// §3.8b — "restore is fail-closed and never silent". Every module that ran
// M_RestoreStationCfg and found an unrecognized image is holding one report;
// this takes them and annunciates each with the OWNING module's canonical path,
// which is what makes the message actionable instead of "something was lost".
//
// The event is AUTO_RESET and therefore never blocking: the consequence belongs
// to E_ConfigRestorePolicy, evaluated in ReleaseReportStart, so a station that
// declared DEFAULTS_AND_ANNUNCIATE really does run while the annunciation
// stands. It stays open until an ENGINEER acknowledges it, because nothing
// makes a lost image come back and an event that closed itself would be a lie.
METHOD PRIVATE _M_DrainRestoreLoss
VAR
    guard    : INT;
    path     : STRING(80);
    expected : UINT;
    found    : UINT;
END_VAR
// §7.7(c) - the local user table is retained outside the module walk; its loss
// is announced and acknowledged exactly like a module's.
IF Access.M_TakeRestoreLoss() THEN
    path := CONCAT(_name, '.Access');
    _M_AnnounceRestoreLoss(Path := path, Text := 'std.error.accessRestoreLost');
END_IF
// Bounded per scan (§5.6): losses are one-shot, so a large subtree simply
// finishes draining over the next few scans instead of stretching one.
FOR guard := 1 TO PL_Fraktal.MAX_EM_CHILDREN DO
    IF NOT M_TakeRestoreLoss(Path => path, Expected => expected, Found => found) THEN
        RETURN;
    END_IF
    _M_AnnounceRestoreLoss(Path := path, Text := 'std.error.configRestoreLost');
END_FOR
END_METHOD

// §3.8b - publish one lost image and open (or extend) its annunciation.
METHOD PRIVATE _M_AnnounceRestoreLoss
VAR_INPUT
    Path : STRING(80);
    Text : STRING(80);
END_VAR
ConfigPersist.RestoreLost := TRUE;
ConfigPersist.RestoreAcknowledged := FALSE;
ConfigPersist.LostPath := Path;
IF _restoreEvt = 0 THEN
    _restoreEvt := AlarmLog.Raise(Reason := E_Reason.CONFIG_RESTORE_LOST,
        Text := Text, Source := Path,
        Severity := E_Severity.MED, Category := E_Category.SYSTEM,
        ResetClass := E_ResetClass.AUTO_RESET);
ELSE
    // A second losing owner gets its own ring entry: a summary that named only
    // the first would hide the rest of the damage.
    _M_RaiseMaintenance(Reason := E_Reason.CONFIG_RESTORE_LOST, Text := Text);
END_IF
END_METHOD

// §3.8b — an operator of at least ENGINEER level accepts that a configuration
// image was lost. Under BLOCK_UNTIL_ACKNOWLEDGED this is what releases
// START_STOP again; under DEFAULTS_AND_ANNUNCIATE it is what clears the
// standing annunciation.
//
// The level is checked directly rather than through a gated action, because
// §3.8b names ENGINEER specifically and a station may legitimately have left
// DATA_WRITE or CONFIG_SET open to a lower level. Acknowledging a lost
// commissioning is a different decision from editing a value.
METHOD AcknowledgeConfigRestore : BOOL
AcknowledgeConfigRestore := FALSE;
IF Access.CurrentLevel < E_AccessLevel.ENGINEER THEN
    RETURN;
END_IF
IF NOT ConfigPersist.RestoreLost THEN
    RETURN;                                // nothing to acknowledge
END_IF
ConfigPersist.RestoreAcknowledged := TRUE;
IF _restoreEvt > 0 THEN
    AlarmLog.Gone(Slot := _restoreEvt);
    _restoreEvt := 0;
END_IF
Access.RecordActivity();
AcknowledgeConfigRestore := TRUE;
END_METHOD

// §3.8b — refuse a set operation, naming the offending record. "One rejection
// aborts the whole load naming the offending (Scope, WriteKey)": a refusal that
// says only "rejected" leaves an engineer diffing two machines by hand.
METHOD PRIVATE _M_RejectConfigSet
VAR_INPUT
    Scope : STRING(80);
    Key   : STRING(160);
END_VAR
ConfigPersist.LastRejectScope := Scope;
ConfigPersist.LastRejectKey := Key;
_M_RaiseMaintenance(Reason := E_Reason.CONFIG_SET_REJECTED,
    Text := 'std.error.configSetRejected');
END_METHOD

// §3.8b — the gate every set operation shares: CONFIG_SET (never DATA_WRITE —
// replacing a machine's entire parametrization is not the same decision as
// changing one number), a wired store, and the owning root READY.
METHOD PRIVATE _M_SetOpAllowed : BOOL
_M_SetOpAllowed := FALSE;
IF NOT _M_ConfigRestored() THEN
    RETURN;
END_IF
IF NOT Access.PermitsLogged(Gate := E_GatedAction.CONFIG_SET) THEN
    RETURN;
END_IF
IF _configStore = 0 THEN
    RETURN;
END_IF
IF _exec <> E_ExecState.READY THEN
    RETURN;
END_IF
_M_SetOpAllowed := TRUE;
END_METHOD

// §3.8b - remove a named set. Gated exactly like save and load (CONFIG_SET, a
// wired store, the root READY) because removing somebody's commissioned set is
// the same order of decision as replacing it, and audited with the set name.
// A store that has held MAX_CONFIG_SETS names needs this to hold a new one.
METHOD DeleteConfigSet : BOOL
VAR_INPUT
    SetName : STRING(80);
END_VAR
DeleteConfigSet := FALSE;
ConfigPersist.LastSetName := SetName;
ConfigPersist.LastSetRecords := 0;
IF NOT _M_SetOpAllowed() THEN
    RETURN;
END_IF
IF NOT _configStore.M_Delete(SetName := SetName) THEN
    RETURN;
END_IF
DeleteConfigSet := TRUE;
// The store's retained memory changed; not durable until written out.
_M_MarkPersistPending();
ListConfigSets();                          // the published listing follows
END_METHOD

// §3.8d - the effective level to read or write one registered value, from
// what its owning module declared and this root's policy. The root's own
// framework keys (unit.modePolicy.*) are in the built-in class. An unknown key
// resolves to ADMIN: the write path refuses it anyway, and a level check must
// never be the thing that lets an unknown key through.
METHOD PRIVATE _M_DataLevelOf : E_AccessLevel
VAR_INPUT
    TargetPath : STRING(255);
    WriteKey   : STRING(160);
    ForWrite   : BOOL;
END_VAR
VAR
    grant    : ST_ConfigAccess;
    minLevel : E_AccessLevel;
END_VAR
_M_DataLevelOf := E_AccessLevel.ADMIN;
IF (TargetPath = Status.Name) AND (LEFT(WriteKey, 16) = 'unit.modePolicy.') THEN
    _M_DataLevelOf := Access.M_DataLevel(ClassId := '', MinLevel := E_AccessLevel.NONE,
        ForWrite := ForWrite);
    RETURN;
END_IF
IF NOT M_ConfigAccessOf(Scope := TargetPath, WriteKey := WriteKey, Grant := grant) THEN
    RETURN;
END_IF
IF ForWrite THEN
    minLevel := grant.MinWriteLevel;
ELSE
    minLevel := grant.MinReadLevel;
END_IF
_M_DataLevelOf := Access.M_DataLevel(ClassId := grant.ClassId, MinLevel := minLevel,
    ForWrite := ForWrite);
END_METHOD

// §3.8d - declare a project data class on this root, at Setup. The levels are
// defaults: a class the deployment already edited keeps its persisted levels.
METHOD M_DeclareDataClass : BOOL
VAR_INPUT
    ClassId    : STRING(80);
    LabelKey   : STRING(160);
    ReadLevel  : E_AccessLevel;
    WriteLevel : E_AccessLevel;
END_VAR
M_DeclareDataClass := Access.M_DeclareClass(ClassId := ClassId,
    LabelKey := LabelKey, ReadLevel := ReadLevel, WriteLevel := WriteLevel);
END_METHOD

// §3.8d/§7.7(b) - edit a class's read or write level. The same gate as
// every other policy edit (ACCESS_POLICY), audited through the mailbox.
METHOD SetDataClassLevel : BOOL
VAR_INPUT
    ClassId  : STRING(160);
    Level    : DINT;
    ForWrite : BOOL;
END_VAR
VAR
    levelReq : E_AccessLevel;
END_VAR
SetDataClassLevel := FALSE;
IF NOT Access.PermitsLogged(Gate := E_GatedAction.ACCESS_POLICY) THEN
    RETURN;
END_IF
IF (Level < TO_DINT(E_AccessLevel.NONE)) OR (Level > TO_DINT(E_AccessLevel.ADMIN))
OR (LEN(ClassId) > 40) THEN
    RETURN;
END_IF
levelReq := Level;                          // range-checked above
SetDataClassLevel := Access.M_SetClassLevel(ClassId := ClassId,
    Level := levelReq, ForWrite := ForWrite);
IF SetDataClassLevel THEN
    ConfigRev := ConfigRev + 1;             // every manifest level may have moved
END_IF
END_METHOD

// §3.8e - TRUE when a (Scope, WriteKey) the subtree did not own names a value of
// the line this Unit references: the line is published under this Unit's own
// scope, and its keys alone begin 'line.'.
METHOD PRIVATE _M_IsLineKey : BOOL
VAR_INPUT
    Scope    : STRING(255);
    WriteKey : STRING(160);
END_VAR
_M_IsLineKey := (_pLine <> 0) AND (Scope = Status.Name)
    AND (LEFT(WriteKey, 5) = 'line.');
END_METHOD

// §3.8e - the subtree first; a line key it does not own goes to the line.
METHOD M_ApplyConfigWrite : BOOL
VAR_INPUT
    Scope     : STRING(255);
    WriteKey  : STRING(160);
    Revision  : UDINT;
    TextValue : STRING(255);
    RootReady : BOOL;
END_VAR
M_ApplyConfigWrite := SUPER^.M_ApplyConfigWrite(Scope := Scope,
    WriteKey := WriteKey, Revision := Revision, TextValue := TextValue,
    RootReady := RootReady);
IF (NOT M_ApplyConfigWrite) AND _M_IsLineKey(Scope := Scope, WriteKey := WriteKey) THEN
    M_ApplyConfigWrite := _pLine^.M_ApplyConfigWrite(Scope := _pLine^.Status.Name,
        WriteKey := WriteKey, Revision := Revision, TextValue := TextValue,
        RootReady := RootReady);
END_IF
END_METHOD

// §3.8e - the staging walk is the write walk, line leg included.
METHOD M_StageConfigWrite : BOOL
VAR_INPUT
    Scope     : STRING(255);
    WriteKey  : STRING(160);
    Revision  : UDINT;
    TextValue : STRING(255);
    RootReady : BOOL;
END_VAR
M_StageConfigWrite := SUPER^.M_StageConfigWrite(Scope := Scope,
    WriteKey := WriteKey, Revision := Revision, TextValue := TextValue,
    RootReady := RootReady);
IF (NOT M_StageConfigWrite) AND _M_IsLineKey(Scope := Scope, WriteKey := WriteKey) THEN
    M_StageConfigWrite := _pLine^.M_StageConfigWrite(Scope := _pLine^.Status.Name,
        WriteKey := WriteKey, Revision := Revision, TextValue := TextValue,
        RootReady := RootReady);
END_IF
END_METHOD

// §3.8e - the capture walk is the write walk, line leg included.
METHOD M_ApplyCapture : BOOL
VAR_INPUT
    Scope     : STRING(255);
    WriteKey  : STRING(160);
    Revision  : UDINT;
    RootReady : BOOL;
END_VAR
M_ApplyCapture := SUPER^.M_ApplyCapture(Scope := Scope, WriteKey := WriteKey,
    Revision := Revision, RootReady := RootReady);
IF (NOT M_ApplyCapture) AND _M_IsLineKey(Scope := Scope, WriteKey := WriteKey) THEN
    M_ApplyCapture := _pLine^.M_ApplyCapture(Scope := _pLine^.Status.Name,
        WriteKey := WriteKey, Revision := Revision, RootReady := RootReady);
END_IF
END_METHOD

// §3.8e/§3.8d - the access walk is the write walk, line leg included, so a line
// value is checked against the level the line declared for it.
METHOD M_ConfigAccessOf : BOOL
VAR_INPUT
    Scope    : STRING(255);
    WriteKey : STRING(160);
END_VAR
VAR_IN_OUT
    Grant : ST_ConfigAccess;
END_VAR
M_ConfigAccessOf := SUPER^.M_ConfigAccessOf(Scope := Scope, WriteKey := WriteKey,
    Grant := Grant);
IF (NOT M_ConfigAccessOf) AND _M_IsLineKey(Scope := Scope, WriteKey := WriteKey) THEN
    M_ConfigAccessOf := _pLine^.M_ConfigAccessOf(Scope := _pLine^.Status.Name,
        WriteKey := WriteKey, Grant := Grant);
END_IF
END_METHOD

// Core §3.8a - declare this root's own recipe record (its ParCfg) and the
// provider it is loaded from. The PAR_CFG values registered inside it become
// editable for EVERY model the root offers (AvailableModels), not only the
// active one, and an edit is written back to the provider's record so a
// changeover keeps it - when the provider is also an I_RecipeStore.
METHOD M_RegisterModelData : BOOL
VAR_INPUT
    pData     : PVOID;
    Size      : UDINT;
    RecipeKey : STRING(80);
    Provider  : I_RecipeProvider;
END_VAR
M_RegisterModelData := FALSE;
IF (pData = 0) OR (Size = 0) OR (Size > PL_Fraktal.MAX_MODEL_DATA_BYTES)
OR (RecipeKey = '') OR (Provider = 0) THEN
    RETURN;
END_IF
_modelProvider := Provider;
__QUERYINTERFACE(Provider, _modelCatalog);
_modelKey := RecipeKey;
M_RegisterModelData := _M_SetModelRegion(pRegion := pData, Size := Size);
END_METHOD

// Serve model-scoped values of AvailableModels[Index] for this one request. 0,
// or the active model's index, is the live record and opens nothing. The record
// is loaded over a copy of the live one, so the provider's SchemaVersion check
// compares like with like. FALSE = no such model, or its record did not load.
METHOD PRIVATE _M_OpenModelView : BOOL
VAR_INPUT
    Index : UDINT;
END_VAR
_M_OpenModelView := FALSE;
_pModelView := 0;
_viewModelCode := '';
IF Index = 0 THEN
    _M_OpenModelView := TRUE;
    RETURN;
END_IF
IF (_modelProvider = 0) OR (_pModelRegion = 0)
OR (Index > TO_UDINT(AvailableModelCount)) THEN
    RETURN;
END_IF
IF AvailableModels[Index].ModelCode = Model.ModelCode THEN
    _M_OpenModelView := TRUE;              // the active model: its record is live
    RETURN;
END_IF
MEMCPY(destAddr := ADR(_modelBuf), srcAddr := _pModelRegion, n := _modelRegionSize);
IF NOT _modelProvider.Load(ModelCode := AvailableModels[Index].ModelCode,
        RecipeKey := _modelKey, pParCfg := ADR(_modelBuf), Size := _modelRegionSize) THEN
    RETURN;
END_IF
_viewModelCode := AvailableModels[Index].ModelCode;
_pModelView := ADR(_modelBuf);
_M_OpenModelView := TRUE;
END_METHOD

// §3.8a - WriteConfig for the model AvailableModels[ModelIndex] (0 = the active
// model). A model-data value is stored in that model's record and saved back to
// the provider; any other value is written as WriteConfig writes it.
METHOD WriteModelConfig : BOOL
VAR_INPUT
    ModelIndex : UDINT;
    TargetPath : STRING(255);
    WriteKey   : STRING(160);
    Revision   : DINT;
    TextValue  : STRING(255);
END_VAR
WriteModelConfig := FALSE;
IF NOT _M_OpenModelView(Index := ModelIndex) THEN
    RETURN;
END_IF
WriteModelConfig := WriteConfig(TargetPath := TargetPath, WriteKey := WriteKey,
    Revision := Revision, TextValue := TextValue);
_pModelView := 0;
END_METHOD

// §3.8a - the manifest walk (M_AppendConfig) with the model-data values of
// AvailableModels[ModelIndex] (0 = the active model). FALSE = no such model.
// For another model the walk yields that model's data only: the rest of the
// manifest is the running station's and is served by index 0.
METHOD M_AppendModelConfig : BOOL
VAR_INPUT
    Pager      : REFERENCE TO FB_ConfigPager;
    ModelIndex : UDINT;
END_VAR
M_AppendModelConfig := FALSE;
IF NOT _M_OpenModelView(Index := ModelIndex) THEN
    RETURN;
END_IF
Pager.M_SetModelOnly(Enabled := ModelIndex > 0);
M_AppendConfig(Pager := Pager);
Pager.M_SetModelOnly(Enabled := FALSE);
_pModelView := 0;
M_AppendModelConfig := TRUE;
END_METHOD

// Write the record a model-scoped value was just stored into back to the
// provider: the viewed model's buffer, or the live record for the active model.
METHOD PRIVATE _M_SaveModelData : BOOL
VAR
    store : I_RecipeStore;
END_VAR
_M_SaveModelData := FALSE;
IF _modelProvider = 0 THEN
    RETURN;
END_IF
IF NOT __QUERYINTERFACE(_modelProvider, store) THEN
    RETURN;
END_IF
IF _pModelView <> 0 THEN
    _M_SaveModelData := store.Save(ModelCode := _viewModelCode, RecipeKey := _modelKey,
        pData := _pModelView, Size := _modelRegionSize);
ELSE
    _M_SaveModelData := store.Save(ModelCode := Model.ModelCode, RecipeKey := _modelKey,
        pData := _pModelRegion, Size := _modelRegionSize);
END_IF
END_METHOD

// §3.8e/§8.5.2 - reference the line this root belongs to (owner or mirror, on
// this controller). A Unit references at most one line; 0 detaches it.
METHOD SetLine : BOOL
VAR_INPUT
    pLine : POINTER TO FB_LineData;
END_VAR
_pLine := pLine;
_lineHost := FALSE;
IF pLine <> 0 THEN
    // The first root to reference a line hosts it (ticks it, lends its log); a
    // line is never a child, so nothing else would run it (§3.8e(a)).
    _lineHost := pLine^.M_BindHost(pHost := THIS, pAlarmLog := ADR(AlarmLog));
END_IF
_shiftInit := FALSE;
CurrentShift := 0;
SetLine := (pLine <> 0);
END_METHOD

// Evaluate only at a finite boundary, or after an empty-calendar edit.
METHOD M_ShiftTick : BOOL
VAR_INPUT
    Now : DT;
    Synchronized : BOOL;
END_VAR
VAR
    idx : INT;
    started : DT;
    ending : DT;
    target : UDINT;
    crossed : BOOL;
    quality : BOOL;
END_VAR
M_ShiftTick := FALSE;
IF _pLine = 0 THEN CurrentShift := 0; ShiftProductionTarget := 0; RETURN; END_IF
IF _shiftInit THEN
    IF Now < _shiftLastNow THEN _shiftSync := FALSE; END_IF
    _shiftLastNow := Now;
    IF (_shiftEnd <> DT#1970-01-01-00:00:00) AND (Now < _shiftEnd) THEN RETURN; END_IF
    IF Now < ShiftStartedAt THEN RETURN; END_IF // no negative history after a backward jump
    IF (_shiftEnd = DT#1970-01-01-00:00:00)
    AND (_shiftCalendarRev = _pLine^.OutImm.Revision) THEN RETURN; END_IF
END_IF
IF NOT _pLine^.M_ShiftInterval(Now := Now, ShiftIndex => idx,
        StartAt => started, EndAt => ending, Target => target) THEN
    _shiftSync := FALSE; RETURN;
END_IF
crossed := _shiftInit AND (_shiftEnd <> DT#1970-01-01-00:00:00);
IF _shiftInit AND NOT crossed AND (idx = 0) THEN
    // Empty/off interval continues; an edit must not erase accrued production.
    _shiftEnd := ending;
    _shiftCalendarRev := _pLine^.OutImm.Revision;
    RETURN;
END_IF
IF _shiftInit THEN
    quality := Synchronized;
    IF crossed AND (DT_TO_UDINT(Now) > DT_TO_UDINT(_shiftEnd) + 1) THEN quality := FALSE; END_IF
    _M_CloseShift(Now := Now, Synchronized := quality);
    M_ShiftTick := TRUE;
END_IF
_shiftInit := TRUE;
CurrentShift := idx;
ShiftStartedAt := Now; // observed start, never invent production before attachment/jump
ShiftProductionTarget := target;
_shiftEnd := ending;
_shiftLastNow := Now;
_shiftCalendarRev := _pLine^.OutImm.Revision;
_shiftSync := Synchronized;
_shiftManualReset := FALSE;
END_METHOD

// §8.5.2(b) - one operation in one scan: record the ending shift as its figures stood,
// then reset the per-shift counts and OEE accumulators (the trend ring is kept). A
// boundary on an unsynchronized clock still closes - stopping the accounting would
// lose more than a late boundary does - and the record says so.
METHOD PRIVATE _M_CloseShift
VAR_INPUT
    Now          : DT;
    Synchronized : BOOL;
END_VAR
VAR
    i         : INT;
    auditSlot : INT;
END_VAR
_M_OeeCompute(); // capture current factors before counters are cleared
FOR i := PL_Fraktal.MAX_SHIFT_HISTORY TO 2 BY -1 DO
    ShiftHistory[i] := ShiftHistory[i - 1];
END_FOR
IF ShiftHistoryCount >= PL_Fraktal.MAX_SHIFT_HISTORY THEN
    ShiftHistoryTruncated := TRUE;
ELSE
    ShiftHistoryCount := ShiftHistoryCount + 1;
END_IF
ShiftHistory[1].SchemaVersion := 3;
ShiftHistory[1].ProductionTarget := ShiftProductionTarget;
ShiftHistory[1].ShiftIndex := CurrentShift;
ShiftHistory[1].StartAt := ShiftStartedAt;
ShiftHistory[1].EndAt := Now;
ShiftHistory[1].TimeSynchronized := _shiftSync AND Synchronized;
ShiftHistory[1].ManualReset := _shiftManualReset;
ShiftHistory[1].GoodCount := GoodCount;
ShiftHistory[1].NokCount := NokCount;
ShiftHistory[1].ReworkCount := ReworkCount;
ShiftHistory[1].RunMs := Oee.RunMs;
ShiftHistory[1].DownMs := Oee.DownMs;
ShiftHistory[1].IdleMs := Oee.IdleMs;
ShiftHistory[1].Availability := Oee.Availability;
ShiftHistory[1].AvailValid := Oee.AvailValid;
ShiftHistory[1].Performance := Oee.Performance;
ShiftHistory[1].PerfValid := Oee.PerfValid;
ShiftHistory[1].Quality := Oee.Quality;
ShiftHistory[1].QualValid := Oee.QualValid;
ShiftHistory[1].Oee := Oee.Oee;
ShiftHistory[1].OeeValid := Oee.OeeValid;
_oeeGoodBase := 0;
_oeeNokBase := 0;
GoodCount := 0;
NokCount := 0;
ReworkCount := 0;
Oee.RunMs := 0;
Oee.DownMs := 0;
Oee.IdleMs := 0;
_M_OeeCompute();
auditSlot := AlarmLog.Raise(Reason := E_Reason.NONE, Text := 'std.audit.shiftClosed',
    Source := _name, Severity := E_Severity.LOW, Category := E_Category.SYSTEM,
    ResetClass := E_ResetClass.AUTO_RESET);
IF auditSlot > 0 THEN
    AlarmLog.Gone(Slot := auditSlot);    // come+gone: into the ring and the event sink
END_IF
END_METHOD

// §3.8b — save the current parametrization as a named set.
//
// The set is a PROJECTION of the same deterministic walk that builds the
// §3.10.2 manifest: M_AppendConfig runs exactly as a QUERY_CONFIG would run it,
// and the pager files every capability of the requested ConfigKind as a
// (Scope, WriteKey) record. There is no second enumeration of "what this
// station's configuration consists of" to drift from the first (§1.1 O9).
//
// Kind selects which of the two kinds of set this is: STATION_CFG for a station
// set (deployment data), PAR_CFG for a model set (one model's recipe data).
METHOD SaveConfigSet : BOOL
VAR_INPUT
    SetName : STRING(80);
    Kind    : E_ConfigKind;
END_VAR
VAR
    info    : ST_ConfigSetInfo;
    records : INT;
END_VAR
SaveConfigSet := FALSE;
ConfigPersist.LastSetName := SetName;
ConfigPersist.LastSetRecords := 0;
IF NOT _M_SetOpAllowed() THEN
    RETURN;
END_IF
IF SetName = '' THEN
    RETURN;
END_IF
info.Used := TRUE;
info.SetName := SetName;
info.RootIdentity := Status.Name;
info.SetSchema := CONFIG_SET_SCHEMA;
info.ConfigRev := ConfigRev;
info.Kind := Kind;
IF Kind = E_ConfigKind.PAR_CFG THEN
    info.ModelCode := Model.ModelCode;     // a model set belongs to ONE model
ELSE
    info.ModelCode := '';
END_IF
info.RecordCount := 0;
info.CreatedAt := F_Now();
info.TimeSynchronized := F_TimeSynchronized();
IF NOT _configPager.M_SetupSetSave(Store := _configStore, Info := info) THEN
    RETURN;
END_IF
M_AppendConfig(Pager := _configPager);     // the SAME walk as the manifest
SaveConfigSet := _configPager.M_FinishSetSave(Records => records);
ConfigPersist.LastSetRecords := records;
IF SaveConfigSet THEN
    // The set now lives in the store's retained memory, which is not durable
    // until it is written out - the same promise as any other accepted write.
    _M_MarkPersistPending();
END_IF
END_METHOD

// §3.8b — apply a named set. STAGED and ALL-OR-NOTHING.
//
// Pass 1 validates every record through its owning module's typed handler and
// changes nothing. Only if all of them pass does pass 2 apply them. A
// half-applied machine parametrization is never a valid outcome, and the only
// way to guarantee that is to know the answer for every record before touching
// the first one.
//
// A record whose capability no longer exists fails pass 1 like any other and is
// REPORTED by name - never silently dropped, because a set that quietly skipped
// the one value that mattered restores a machine to almost its commissioned
// state, which is the failure that is hardest to notice.
METHOD LoadConfigSet : BOOL
VAR_INPUT
    SetName : STRING(80);
END_VAR
VAR
    info    : ST_ConfigSetInfo;
END_VAR
LoadConfigSet := FALSE;
ConfigPersist.LastSetName := SetName;
ConfigPersist.LastSetRecords := 0;
ConfigPersist.LastRejectScope := '';
ConfigPersist.LastRejectKey := '';
IF NOT _M_SetOpAllowed() THEN
    RETURN;
END_IF
IF NOT _M_CopySet(SetName := SetName) THEN
    RETURN;
END_IF
IF NOT _loadSnapshot.M_ReadInfo(SetName := SetName, Info := info) THEN
    _M_RejectConfigSet(Scope := '', Key := SetName);
    RETURN;
END_IF
IF info.RootIdentity <> Status.Name THEN
    // The set carries the identity of the root that produced it precisely so
    // this can be asked. Every record's Scope is prefixed by that identity, so
    // a mismatch would fail record by record anyway - naming the root instead
    // tells the operator WHY in one line.
    _M_RejectConfigSet(Scope := info.RootIdentity, Key := '');
    RETURN;
END_IF
IF info.Kind = E_ConfigKind.PAR_CFG THEN
    // §3.8b: a MODEL set "shall be applied through the §3.8 changeover
    // transaction (PrepareRecipe -> recursive readiness -> infallible
    // CommitRecipe), never as a sequence of per-field writes". Applying it here
    // would be exactly that forbidden sequence, so it is refused. Saving a
    // model set is supported; loading one is a changeover this build does not
    // implement, and refusing is the honest half of that.
    _M_RejectConfigSet(Scope := info.ModelCode, Key := '');
    RETURN;
END_IF
IF NOT _M_CaptureConfig(SetName := '_validation', Kind := info.Kind, ModelIndex := 0) THEN RETURN; END_IF
IF NOT _M_ValidateSetShape(Store := _loadSnapshot, Info := info, AnyRevision := FALSE) THEN
    RETURN;
END_IF
IF NOT _M_ApplySet(SetName := SetName, RecordCount := info.RecordCount, Kind := info.Kind,
        Restoring := FALSE) THEN
    RETURN;
END_IF
ConfigRev := ConfigRev + 1;
ConfigPersist.LastSetRecords := info.RecordCount;
_M_MarkPersistPending();
_M_RaiseMaintenance(Reason := E_Reason.EVENT_CONFIG_SET_APPLIED,
    Text := 'std.audit.configSetApplied');
LoadConfigSet := TRUE;
END_METHOD

// §3.8b - replay the set frozen in _loadSnapshot. STAGED and ALL-OR-NOTHING:
// pass 1 validates every record through its owning module's typed handler and
// changes nothing; only if all of them pass does pass 2 apply them. A record
// whose capability no longer exists fails pass 1 like any other and is named.
//
// Shared by an operator's LoadConfigSet and the start-up restore of the live
// documents. Restoring skips the session's per-value level (§3.8d(e)): those
// values were accepted once already, and replaying them is the machine's act,
// not an operator's. With a model view open the values go to that record.
METHOD PRIVATE _M_ApplySet : BOOL
VAR_INPUT
    SetName     : STRING(80);
    RecordCount : INT;
    Kind        : E_ConfigKind;
    Restoring   : BOOL;
END_VAR
VAR
    record    : ST_ConfigRecord;
    i         : INT;
    applied   : BOOL;
    lineBatch : BOOL;
END_VAR
_M_ApplySet := FALSE;
lineBatch := (Kind = E_ConfigKind.LINE_CFG) AND (_pLine <> 0);
IF lineBatch THEN
    IF NOT _pLine^.M_BeginConfigBatch() THEN RETURN; END_IF
END_IF
// ---- pass 1: stage. Nothing in the machine changes in this loop. ----
FOR i := 1 TO RecordCount DO
    IF NOT _loadSnapshot.M_ReadRecord(SetName := SetName, Index := i,
            Record := record) THEN
        _M_RejectConfigSet(Scope := '', Key := SetName);
        IF lineBatch THEN _pLine^.M_EndConfigBatch(); END_IF
        RETURN;
    END_IF
    // §3.8d(e) - CONFIG_SET alone cannot replace a value this session could
    // not edit one at a time. Checked in the staging pass, so nothing moved.
    IF NOT Restoring THEN
        IF NOT Access.M_PermitsLevelLogged(Required := _M_DataLevelOf(TargetPath := record.Scope,
                WriteKey := record.WriteKey, ForWrite := TRUE)) THEN
            _M_RejectConfigSet(Scope := record.Scope, Key := record.WriteKey);
            IF lineBatch THEN _pLine^.M_EndConfigBatch(); END_IF
            RETURN;
        END_IF
    END_IF
    IF NOT _M_StageOneRecord(Record := record) THEN
        _M_RejectConfigSet(Scope := record.Scope, Key := record.WriteKey);
        IF lineBatch THEN _pLine^.M_EndConfigBatch(); END_IF
        RETURN;
    END_IF
END_FOR
IF lineBatch THEN
    IF NOT _pLine^.M_ValidateConfigBatch() THEN
        _pLine^.M_EndConfigBatch(); _M_RejectConfigSet(Scope := Status.Name, Key := SetName); RETURN;
    END_IF
END_IF
// ---- pass 2: apply. Every record already proved acceptable on the SAME
// validator, so a refusal here cannot be a data problem. ----
FOR i := 1 TO RecordCount DO
    IF NOT _loadSnapshot.M_ReadRecord(SetName := SetName, Index := i,
            Record := record) THEN
        IF lineBatch THEN _pLine^.M_EndConfigBatch(); END_IF
        _M_ConfigSetHalfApplied(Scope := record.Scope, Key := record.WriteKey);
        RETURN;
    END_IF
    applied := _M_WriteBaseConfig(TargetPath := record.Scope,
        WriteKey := record.WriteKey, Revision := record.Revision,
        TextValue := record.ValueText, Commit := TRUE);
    IF NOT applied THEN
        applied := M_ApplyConfigWrite(Scope := record.Scope,
            WriteKey := record.WriteKey, Revision := record.Revision,
            TextValue := record.ValueText,
            RootReady := (_exec = E_ExecState.READY) OR (_pModelView <> 0));
    END_IF
    IF NOT applied THEN
        IF lineBatch THEN _pLine^.M_EndConfigBatch(); END_IF
        _M_ConfigSetHalfApplied(Scope := record.Scope, Key := record.WriteKey);
        RETURN;
    END_IF
END_FOR
IF lineBatch THEN
    _pLine^.M_CommitConfigBatch();
END_IF
_M_ApplySet := TRUE;
END_METHOD

// §3.8b — would this record be accepted? The same two-step the write path
// takes: framework-owned keys first, then the recursive walk to the owning
// module. Sharing the writers' own code with Commit := FALSE is what makes
// "staged" mean something: a separate validator could pass a record the write
// path would then refuse, and the load would be half-applied after all.
METHOD PRIVATE _M_StageOneRecord : BOOL
VAR_INPUT
    Record : ST_ConfigRecord;
END_VAR
_M_StageOneRecord := _M_WriteBaseConfig(TargetPath := Record.Scope,
    WriteKey := Record.WriteKey, Revision := Record.Revision,
    TextValue := Record.ValueText, Commit := FALSE);
IF _M_StageOneRecord THEN
    RETURN;
END_IF
_M_StageOneRecord := M_StageConfigWrite(Scope := Record.Scope,
    WriteKey := Record.WriteKey, Revision := Record.Revision,
    TextValue := Record.ValueText,
    // Another model's record is not what the machine is running on.
    RootReady := (_exec = E_ExecState.READY) OR (_pModelView <> 0));
END_METHOD

// §3.8b — a record passed staging and then failed to apply. This cannot
// happen: both run the same validator on the same data in the same scan. If it
// ever does, the machine is half-parametrized and that is a state the standard
// says is never valid - so it is escalated as a BLOCKING alarm rather than
// returned as a FALSE somebody might retry. A framework defect that leaves a
// machine half-configured has to stop it, not inconvenience it.
METHOD PRIVATE _M_ConfigSetHalfApplied
VAR_INPUT
    Scope : STRING(80);
    Key   : STRING(160);
END_VAR
ConfigPersist.LastRejectScope := Scope;
ConfigPersist.LastRejectKey := Key;
AlarmLog.Raise(Reason := E_Reason.CONFIG_SET_REJECTED,
    Text := 'std.error.configSetHalfApplied', Source := Scope,
    Severity := E_Severity.HIGH, Category := E_Category.SYSTEM,
    ResetClass := E_ResetClass.MANUAL_RESET);
END_METHOD

// §3.8b — refresh the published listing of stored sets. Read-only, so it is
// gated on CONFIG_SET without the audited write path: seeing which sets exist
// is not replacing a machine's parametrization.
METHOD ListConfigSets : BOOL
VAR
    i     : INT;
    total : INT;
END_VAR
ListConfigSets := FALSE;
FOR i := 1 TO PL_Fraktal.MAX_CONFIG_SETS DO
    ConfigSets[i].Used := FALSE;
    ConfigSets[i].SetName := '';
    ConfigSets[i].RecordCount := 0;
END_FOR
ConfigSetCount := 0;
IF NOT Access.Permits(Gate := E_GatedAction.CONFIG_SET) THEN
    RETURN;
END_IF
IF _configStore = 0 THEN
    RETURN;
END_IF
total := _configStore.M_Count();
FOR i := 1 TO PL_Fraktal.MAX_CONFIG_SETS DO
    IF i > total THEN
        EXIT;
    END_IF
    IF _configStore.M_InfoAt(Index := i, Info := ConfigSets[i]) THEN
        ConfigSetCount := i;
    END_IF
END_FOR
ListConfigSets := TRUE;
END_METHOD

// §3.8b — serve one line of a set's JSON document. Line 0 is the header and
// 1..RecordCount are the records, so a client pulls a movable document a line
// at a time and no full document buffer ever exists in the PLC - the same
// paging discipline QUERY_CONFIG already uses for the manifest.
//
// This is what makes a set MOVABLE, which is the point of naming sets at all: a
// station's commissioning can leave the controller as text, be reviewed,
// diffed, version-controlled and put on the next machine.
METHOD ExportConfigSetLine : BOOL
VAR_INPUT
    SetName : STRING(80);
    Line    : INT;
END_VAR
VAR
    info   : ST_ConfigSetInfo;
    record : ST_ConfigRecord;
END_VAR
ExportConfigSetLine := FALSE;
ConfigSetDocument := '';
ConfigSetDocumentLine := Line;
ConfigSetDocumentLines := 0;
IF NOT Access.Permits(Gate := E_GatedAction.CONFIG_SET) THEN
    RETURN;
END_IF
IF _configStore = 0 THEN
    RETURN;
END_IF
IF NOT _configStore.M_ReadInfo(SetName := SetName, Info := info) THEN
    RETURN;
END_IF
ConfigSetDocumentLines := info.RecordCount;
IF Line <= 0 THEN
    ConfigSetDocument := _setJson.M_Header(Info := info);
ELSE
    IF NOT _configStore.M_ReadRecord(SetName := SetName, Index := Line,
            Record := record) THEN
        RETURN;
    END_IF
    IF NOT Access.M_PermitsLevel(Required := _M_DataLevelOf(TargetPath := record.Scope,
            WriteKey := record.WriteKey, ForWrite := FALSE)) THEN
        RETURN;                           // §3.8d(e): the export fails, it is not thinned
    END_IF
    ConfigSetDocument := _setJson.M_Record(Record := record);
END_IF
// An empty line means the projection REFUSED to render it rather than shorten
// it, so the export fails here instead of shipping a document with a hole.
ExportConfigSetLine := (ConfigSetDocument <> '');
END_METHOD

// §3.8b — take one line of a set's JSON document back in. A header line opens
// a store save, record lines append to it, and Commit closes it.
//
// Import writes into the STORE, never into the machine. Bringing a document in
// and applying it to the equipment are two decisions, and keeping them apart is
// what lets LoadConfigSet stay staged and all-or-nothing: an imported set is
// validated against THIS machine's capabilities when somebody chooses to load
// it, not silently as it arrives.
//
// Everything here is untrusted input in the fullest sense - hand-edited, from
// another vendor's tool, from another machine - so the line is parsed into a
// typed record and nothing more is assumed about it (§5.6, §14).
METHOD ImportConfigSetLine : BOOL
VAR_INPUT
    Line   : STRING(480);
    Commit : BOOL;
END_VAR
VAR
    info   : ST_ConfigSetInfo;
    record : ST_ConfigRecord;
END_VAR
ImportConfigSetLine := FALSE;
IF NOT _M_SetOpAllowed() THEN
    _importOpen := FALSE;
    RETURN;
END_IF
IF _setJson.M_ParseHeader(Line := Line, Info := info) THEN
    _importOpen := FALSE;
    info.Used := TRUE;
    info.RecordCount := 0;
    IF NOT _configStore.M_SaveBegin(Info := info) THEN
        RETURN;
    END_IF
    _importOpen := TRUE;
    ConfigPersist.LastSetName := info.SetName;
    ImportConfigSetLine := TRUE;
    RETURN;
END_IF
IF NOT _importOpen THEN
    RETURN;                                // a record before its header: refuse
END_IF
IF _setJson.M_ParseRecord(Line := Line, Record := record) THEN
    ImportConfigSetLine := _configStore.M_SaveRecord(Record := record);
    IF NOT ImportConfigSetLine THEN
        _configStore.M_SaveAbort();
        _importOpen := FALSE;
        RETURN;
    END_IF
ELSIF NOT Commit THEN
    // Neither a header nor a record, and not the closing call: the document is
    // not one this build understands. Abort rather than commit a partial set.
    _configStore.M_SaveAbort();
    _importOpen := FALSE;
    RETURN;
END_IF
IF Commit THEN
    ImportConfigSetLine := _configStore.M_SaveCommit();
    _importOpen := FALSE;
    IF ImportConfigSetLine THEN
        _M_MarkPersistPending();
    END_IF
END_IF
END_METHOD

// §3.8b - take part of a set line. A request carries at most 255 characters
// and an exported line may hold 480, so a longer line arrives as pieces:
// More = TRUE holds this piece and waits for the next; the first piece without
// More completes the line, which is then imported exactly like a whole one.
//
// Joined by FB_ConfigSetJson.M_Join, which measures first: a line that would
// exceed its width is refused and the import aborted - never truncated. (Not
// CONCAT/LEN: those stop at 255, which is the very limit being crossed.)
METHOD ImportConfigSetPiece : BOOL
VAR_INPUT
    Piece  : STRING(255);
    More   : BOOL;
    Commit : BOOL;
END_VAR
VAR
    line : STRING(480);
END_VAR
ImportConfigSetPiece := FALSE;
IF NOT _M_SetOpAllowed() THEN
    _importPart := '';
    RETURN;
END_IF
line := _importPart;
IF NOT _setJson.M_Join(Tail := Piece, Line := line) THEN
    _importPart := '';
    IF _importOpen THEN
        _configStore.M_SaveAbort();
        _importOpen := FALSE;
    END_IF
    RETURN;
END_IF
IF More THEN
    _importPart := line;
    ImportConfigSetPiece := TRUE;             // held, not yet imported
    RETURN;
END_IF
_importPart := '';
ImportConfigSetPiece := ImportConfigSetLine(Line := line, Commit := Commit);
END_METHOD

METHOD M_SequenceAskDecision
VAR_INPUT
    Req : ST_DecisionRequest;
END_VAR
_M_AskDecision(Req := Req);
END_METHOD

METHOD M_SequenceAwait : BOOL
VAR_INPUT
    Idx : INT;
    Label : STRING(120);
    Ok : BOOL;
END_VAR
M_SequenceAwait := _M_Await(Idx := Idx, Label := Label, Ok := Ok);
END_METHOD

METHOD M_SequenceClearDecision
IF Decision.Prompt <> '' THEN
    _M_LogDecision(EventKey := 'std.audit.decisionWithdrawn',
        SourcePath := Decision.SourcePath, Option := 0);
END_IF
_M_ClearDecisionState();
END_METHOD

METHOD M_SequenceComplete
IF _mode = E_Mode.CHANGEOVER THEN
    _M_HostEvent(Kind := E_HostEventKind.CHANGEOVER_DONE, PartUid := '',
        Subject := 'Model', Value := Model.ModelCode,
        Verdict := E_Verdict.NONE, ReasonCode := E_Reason.NONE);
END_IF
_M_Complete();
END_METHOD

METHOD M_SequenceCountGood
CountGood();
END_METHOD

METHOD M_SequenceEndOfCycle : BOOL
M_SequenceEndOfCycle := _M_EndOfCycle();
END_METHOD

METHOD M_SequenceFault
VAR_INPUT
    Reason : E_Reason;
    DescriptionKey : STRING(255);
END_VAR
_M_Fault(Reason, DescriptionKey);
END_METHOD

METHOD M_SequencePartProcessed : BOOL
VAR_INPUT
    Verdict : E_Verdict;
    Reason : E_Reason;
END_VAR
M_SequencePartProcessed :=
    _M_PartProcessed(Verdict := Verdict, Reason := Reason);
END_METHOD

METHOD M_SequencePartReceived : BOOL
M_SequencePartReceived := _M_PartReceived();
END_METHOD

METHOD M_SequencePartRecord : BOOL
VAR_INPUT
    RecordName : STRING(64);
    Value : LREAL;
    Minimum : LREAL;
    Maximum : LREAL;
    Target : LREAL;
    EngUnit : STRING(16);
END_VAR
M_SequencePartRecord := _M_PartRecord(RecordName := RecordName,
    Value := Value, Minimum := Minimum, Maximum := Maximum, Target := Target,
    EngUnit := EngUnit);
END_METHOD

METHOD M_SequencePartStarted
_M_PartStarted();
END_METHOD

// §6.8 register an attached chain (idempotent, bounded). Called from
// FB_SequenceBase.M_Attach, never by project code.
METHOD M_SequenceRegister : BOOL
VAR_INPUT
    Seq : I_Sequence;
END_VAR
VAR
    i : INT;
END_VAR
M_SequenceRegister := FALSE;
IF Seq = 0 THEN
    RETURN;
END_IF
FOR i := 1 TO _sequenceCount DO
    IF _sequences[i] = Seq THEN
        M_SequenceRegister := TRUE;        // already attached: Setup ran again
        RETURN;
    END_IF
END_FOR
IF _sequenceCount >= PL_Fraktal.MAX_SEQUENCES THEN
    RETURN;                                // bounded; refused, never silently dropped
END_IF
_sequenceCount := _sequenceCount + 1;
_sequences[_sequenceCount] := Seq;
M_SequenceRegister := TRUE;
END_METHOD

// §6.10 — reset every attached chain's shared transition result once per
// PLC cycle, before _M_Dispatch drives any step action. This is why a project
// never calls M_BeginScan itself, and why an SFC/LD/FBD chart needs no wiring
// to be safe against a stale ADVANCE (O1).
METHOD PROTECTED _M_BeginSequenceScan
VAR
    i : INT;
END_VAR
// §6.12 — close out the legs the previous scan's dispatch stopped recording. A step
// is live exactly while its action keeps calling M_Step, which is the same fact the
// chart draws, so nothing has to be deregistered when a leg finishes. Sweeping legs
// rather than rows makes this ~10 iterations however long the chain is.
FOR i := 0 TO PL_Fraktal.MAX_PARALLEL_BRANCHES DO
    IF (ActiveSteps[i].RowIdx > 0) AND NOT _branchTouched[i] THEN
        // The row keeps how long it ran: the HMI polls too slowly to have timed it.
        SequenceSteps[ActiveSteps[i].RowIdx].LastDuration := ActiveSteps[i].Elapsed;
        ActiveSteps[i].RowIdx := 0;
        ActiveSteps[i].TimedOut := FALSE;
    END_IF
    _branchTouched[i] := FALSE;
END_FOR
FOR i := 1 TO _sequenceCount DO
    IF _sequences[i] <> 0 THEN
        _sequences[i].M_BeginScan();
    END_IF
END_FOR
END_METHOD

// §6.8 - restart every attached chain. The base calls it where a chain can never
// resume (first scan, mode change, abort, abort in error). Whether a fresh run
// command or an operator reset RESTARTS the chain or lets it resume where an
// error stopped it is the project's policy (§6.9(d)), so a project that wants a
// restart there calls this one line from OnCommandStart / OnOperatorReset.
METHOD PROTECTED _M_RestartSequences
VAR
    i : INT;
END_VAR
FOR i := 1 TO _sequenceCount DO
    IF _sequences[i] <> 0 THEN
        _sequences[i].M_Restart();
    END_IF
END_FOR
// A decision belongs to the chain step that asked it; a restarted chain asks again.
Decision.Prompt := '';
DecisionAnswer := 0;
END_METHOD

// §3.14 - an aborted mode chain is abandoned, never resumed: restart every
// attached chain so the next command starts at N000 (§6.8).
METHOD PROTECTED OnAbort : DINT
OnAbort := SUPER^.OnAbort();
_M_RestartSequences();
END_METHOD

// §3.14 - error-state abort abandons the chain the same way (§6.8).
METHOD PROTECTED OnAbortInError : DINT
OnAbortInError := SUPER^.OnAbortInError();
_M_RestartSequences();
END_METHOD

// §6.9(e) — a step said something worth recording that is not a failure.
// Deliberately does NOT touch _exec: no fault is adopted, _M_Dispatch keeps
// running, and the chain follows its own recovery path. The ring entry is
// AUTO_RESET come+gone (§8.3(c)) so it can never block the next Start.
METHOD M_SequenceWarn : BOOL
VAR_INPUT
    Diag : ST_Diagnostic;
END_VAR
VAR
    d    : ST_Diagnostic;
    slot : INT;
END_VAR
d := Diag;
IF d.SourcePath = '' THEN
    d.SourcePath := _name;
END_IF
F_RationalizeDiagnostic(Diag := d);   // §8.8 owns a registered reason's level
IF (_seqIndex >= 1) AND (_seqIndex <= SequenceStepCount) THEN
    SequenceSteps[_seqIndex].WarningActive := TRUE;
    // A message about THIS Unit has nowhere to drill; one about a child keeps the
    // child's path, so the chart links to the module the message is about.
    IF d.SourcePath = _name THEN
        _M_SequenceAnnotate(RowIdx := _seqIndex, IsError := FALSE,
            Key := d.Description, SourcePath := '');
    ELSE
        _M_SequenceAnnotate(RowIdx := _seqIndex, IsError := FALSE,
            Key := d.Description, SourcePath := d.SourcePath);
    END_IF
END_IF
slot := AlarmLog.Raise(Reason := d.ReasonCode, Text := d.Description,
    Source := d.SourcePath, Severity := d.Severity, Category := d.Category,
    ResetClass := E_ResetClass.AUTO_RESET);
IF slot > 0 THEN
    AlarmLog.Gone(Slot := slot);       // an occurrence, not a standing condition
END_IF
M_SequenceWarn := TRUE;
END_METHOD

// §6.9 — a step raised a first-out itself. Stamp the flow-chart row with the
// error and its link before adopting the diagnostic, so the §3.13 chart can mark
// the step red and drill into the module that actually failed even when the step
// passed Awaits := 0. Adopting the diagnostic stops the chain: _M_FaultDiag puts
// the Unit in ERROR and _M_Dispatch no longer runs.
METHOD M_SequenceRaise : BOOL
VAR_INPUT
    Diag     : ST_Diagnostic;
    LinkPath : STRING(255);
END_VAR
M_SequenceRaise := FALSE;
IF (_seqIndex >= 1) AND (_seqIndex <= SequenceStepCount) THEN
    SequenceSteps[_seqIndex].ErrorActive := TRUE;
    _M_SequenceAnnotate(RowIdx := _seqIndex, IsError := TRUE,
        Key := Diag.Description, SourcePath := LinkPath);
END_IF
_M_FaultDiag(Diag := Diag);
M_SequenceRaise := TRUE;
END_METHOD

// §6.9 — the ERROR state ended: clear the flow-chart error marks and re-arm
// every attached chain so the step that raised the fault re-evaluates its
// command. A project writes nothing for this (§1.1 O1).
METHOD PROTECTED _M_ResumeSequencesAfterError
VAR
    i : INT;
END_VAR
FOR i := 1 TO SequenceStepCount DO
    SequenceSteps[i].ErrorActive := FALSE;
END_FOR
_M_SequenceAnnotationClear(RowIdx := 0, IsError := TRUE);
FOR i := 1 TO _sequenceCount DO
    IF _sequences[i] <> 0 THEN
        _sequences[i].M_ResumeAfterError();
    END_IF
END_FOR
END_METHOD

// I_SequenceHost (§6.7/§6.8) — step record for a separately-compiled chain.
METHOD M_SequenceSetStep
VAR_INPUT
    StepNo : INT;
    StepName : STRING(120);
    Awaits : I_Module;
    AwaitingLabel : STRING(120);
    TimeClass : E_TimeClass;
    ExpectedTime : TIME;
    Branch : INT;
END_VAR
// §6.12 — a step on a concurrent LEG publishes its own row and nothing else. The
// Unit's CurrentStep, the §6.9 stall walk and the §8.11.4 profiler are singular by
// definition; letting a leg write them would make the walk report whichever leg
// happened to run last. A leg is timed and guarded on its own row instead, so
// _M_SetStep keeps the signature every inline chain already calls (§1.1 O1).
IF Branch > 0 THEN
    _M_RecordSequenceStep(StepNo := StepNo, StepName := StepName, Awaits := Awaits,
        AwaitingLabel := AwaitingLabel, TimeClass := TimeClass, ExpectedTime := ExpectedTime,
        Branch := Branch);
    RETURN;
END_IF
_M_SetStep(StepNo := StepNo, StepName := StepName,
    Awaits := Awaits, AwaitingLabel := AwaitingLabel, TimeClass := TimeClass,
    ExpectedTime := ExpectedTime);
END_METHOD

METHOD M_SequenceStepGate : BOOL
VAR_INPUT
    Steppable : BOOL;
END_VAR
M_SequenceStepGate := _M_StepGate(Steppable := Steppable);
END_METHOD

// §3.4/§8.11 — accept a pending Stop BETWEEN cycles: the open profile fragment
// (just the wait step) is abandoned, not published as a production cycle.
METHOD M_SequenceStopNow
Profiler.CycleAbandon();
_stopReq := FALSE;
Execute := FALSE;
_M_Complete();
END_METHOD

// §3.4 — a chain polls this at its between-cycles wait step.
METHOD M_SequenceStopPending : BOOL
M_SequenceStopPending := _stopReq AND (_exec = E_ExecState.BUSY);
END_METHOD

METHOD M_SequenceTakeDecision : INT
M_SequenceTakeDecision := _M_TakeDecision();
END_METHOD

// §7.6.1a — single gated entry for a HELD manual action (hold-to-run). Same
// gates as ManualCommandTo: this Unit in MANUAL (§3.4) and MANUAL access
// (§7.7). Held := TRUE latches the request; FALSE releases it immediately.
//
// The release is explicit AND the latch expires, deliberately both: an explicit
// release stops the motion the moment the operator lets go, and the deadline
// stops it when no release ever arrives because the client vanished. Relying on
// either alone leaves one of those two cases moving.
//
// Hold-to-run over a transport is NON-SAFETY (no dead-man, TC3 §7.6): the
// enabling device is the safety-rated fact, derived below from the §9 facet and
// carried to the module, which weighs it itself.
METHOD ManualHeldTo : BOOL
VAR_INPUT
    TargetPath : STRING(255);
    Value      : DINT;
    Held       : BOOL;
END_VAR
VAR
    auditSlot : INT;
END_VAR
ManualHeldTo := FALSE;
IF NOT Held THEN
    // A release is always honoured, whatever the mode or access says now. The
    // operator letting go must never depend on a gate that may have changed
    // since they took hold of it.
    _heldActive := FALSE;
    _heldPath := '';
    _heldValue := 0;
    ManualHeldTo := TRUE;
    RETURN;
END_IF
IF _mode <> E_Mode.MANUAL THEN
    auditSlot := AlarmLog.Raise(Reason := E_Reason.NONE,
        Text := 'std.audit.manualCommandWrongMode', Source := TargetPath,
        Severity := E_Severity.LOW, Category := E_Category.SYSTEM,
        ResetClass := E_ResetClass.AUTO_RESET);
    IF auditSlot > 0 THEN AlarmLog.Gone(Slot := auditSlot); END_IF
    RETURN;
END_IF
IF NOT Access.PermitsLogged(Gate := E_GatedAction.MANUAL) THEN
    RETURN;                              // §7.7 denial already audited
END_IF
// Prove the target accepts it BEFORE latching, so a hold on a module that
// refuses never becomes a standing request nobody can see the source of.
IF NOT _M_RouteHeld(TargetPath := TargetPath, Value := Value) THEN
    RETURN;
END_IF
_heldPath := TargetPath;
_heldValue := Value;
_heldActive := TRUE;
_heldSinceMs := TIME_TO_DWORD(TIME());
ManualHeldTo := TRUE;
END_METHOD

// §7.6.1a — derive the enabling-device fact from THIS root's §9 safety facet and
// carry it to the owning module through the registered-child walk.
//
// F_ManualEnable is the single place the fact is derived, so grepping for it
// lists every path by which motion is authorised by an enabling device. Until
// now it had no production caller at all - the capability existed and nothing
// reached it.
METHOD PROTECTED _M_RouteHeld : BOOL
VAR_INPUT
    TargetPath : STRING(255);
    Value      : DINT;
END_VAR
VAR
    enable : ST_ManualEnableStatus;
END_VAR
enable := F_ManualEnable(Safety := Safety);
_M_RouteHeld := M_ApplyHeld(Scope := TargetPath, Value := Value,
    Enable := enable);
END_METHOD

// §3.13/§3.10.2 — raise the manifest revision ONCE the flow chart has stopped
// growing, rather than once per row discovered.
//
// The rows are the manifest's largest and most volatile contributor and they
// appear one at a time as the chain visits them, so a per-row bump turned one
// mode entry into one full-manifest refetch per step. This waits for the burst
// to settle and then charges for it once.
//
// The delay is bounded and small (PL_Fraktal.CHART_REV_SETTLE_MS): the chart
// appears fractionally later and COMPLETE, instead of promptly and then being
// refetched fourteen more times.
METHOD PRIVATE _M_ChartRevCyclic
VAR
    elapsed : DWORD;
END_VAR
IF NOT _chartDirty THEN
    RETURN;
END_IF
// Unsigned subtraction, so the monotonic counter wrapping cannot fabricate a
// settled chart (TC3 §8.11).
elapsed := TIME_TO_DWORD(TIME()) - _chartTouchedMs;
IF elapsed < PL_Fraktal.CHART_REV_SETTLE_MS THEN
    RETURN;                            // still growing: let the burst finish
END_IF
_chartDirty := FALSE;
ConfigRev := ConfigRev + 1;
END_METHOD

// §7.6.1a — re-assert the latched hold every scan, and drop it when the client
// stops refreshing. The module's own freshness timer stops the motion; this
// stops the ROOT from going on asking for it.
METHOD PRIVATE _M_HeldCyclic
VAR
    elapsed : DWORD;
END_VAR
IF NOT _heldActive THEN
    RETURN;
END_IF
// Leaving MANUAL, or losing the access that granted it, ends the hold at once.
IF _mode <> E_Mode.MANUAL THEN
    _heldActive := FALSE;
    RETURN;
END_IF
IF NOT Access.Permits(Gate := E_GatedAction.MANUAL) THEN
    _heldActive := FALSE;
    RETURN;
END_IF
// Unsigned subtraction, so the monotonic counter wrapping cannot fabricate an
// expired hold (TC3 §8.11).
elapsed := TIME_TO_DWORD(TIME()) - _heldSinceMs;
IF elapsed > PL_Fraktal.MANUAL_HELD_REFRESH_MS THEN
    _heldActive := FALSE;                // client went quiet: let go for it
    RETURN;
END_IF
_M_RouteHeld(TargetPath := _heldPath, Value := _heldValue);
END_METHOD

// §7.6.1 — single gated manual-command entry for the HMI. Accepts ONLY when this
// Unit is in MANUAL (§3.4) AND the user holds MANUAL access (§7.7). Routes to the
// target module's ManualCommand (through the command surface — defended, not
// bypassed). Logs every accept/reject as a §8.3 event. Concrete Units override
// _M_RouteManual to map TargetPath -> the child module.
METHOD ManualCommandTo : BOOL
VAR_INPUT
    TargetPath : STRING(255);
    Value : DINT;
END_VAR
VAR
    auditSlot : INT;
END_VAR
ManualCommandTo := FALSE;
IF _mode <> E_Mode.MANUAL THEN
    auditSlot := AlarmLog.Raise(Reason := E_Reason.NONE,
        Text := 'std.audit.manualCommandWrongMode', Source := TargetPath,
        Severity := E_Severity.LOW, Category := E_Category.SYSTEM, ResetClass := E_ResetClass.AUTO_RESET);
    IF auditSlot > 0 THEN AlarmLog.Gone(Slot := auditSlot); END_IF
    RETURN;
END_IF
IF NOT Access.PermitsLogged(Gate := E_GatedAction.MANUAL) THEN
    RETURN;                              // §7.7 denial already audited
END_IF
ManualCommandTo := _M_RouteManual(TargetPath := TargetPath, Value := Value);
IF ManualCommandTo THEN
    auditSlot := AlarmLog.Raise(Reason := E_Reason.NONE,
        Text := 'std.audit.manualCommandAccepted', Source := TargetPath,
        Severity := E_Severity.LOW, Category := E_Category.SYSTEM, ResetClass := E_ResetClass.AUTO_RESET);
ELSE
    auditSlot := AlarmLog.Raise(Reason := E_Reason.UNSUPPORTED_COMMAND,
        Text := 'std.audit.manualCommandRejected', Source := TargetPath,
        Severity := E_Severity.LOW, Category := E_Category.SYSTEM, ResetClass := E_ResetClass.AUTO_RESET);
END_IF
IF auditSlot > 0 THEN AlarmLog.Gone(Slot := auditSlot); END_IF
END_METHOD

PROPERTY ModeActive : E_Mode
GET
ModeActive := _mode;
END_GET
END_PROPERTY

PROPERTY ModelCode : STRING(64)
GET
ModelCode := Model.ModelCode;
END_GET
END_PROPERTY

PROPERTY ModuleType : E_ModuleType
GET
ModuleType := E_ModuleType.UNIT;
END_GET
END_PROPERTY

// base first (§3.14.2); then children, one-shot init, mode transition, stall watch
METHOD PROTECTED OnCyclic : DINT
VAR
    publishIdx : INT;
    modeIdx    : E_Mode;
    styleIdx   : E_RunStyle;
    previousMode : E_Mode;
    modeExitResult : DINT;
    highestSeverity : E_Severity;
    alarmActive : BOOL;
    heldReported : BOOL;
END_VAR
OnCyclic := SUPER^.OnCyclic();
_M_SyncModelCatalog();
_M_BeginSequenceScan();                               // §6.10 one-scan result reset for every attached chain
_M_TickChildren();
IF _pLine <> 0 THEN
    IF _lineHost THEN
        _pLine^.Cyclic();                             // §3.8e the hosting root runs the line
    END_IF
    // A line value can change without a write through THIS root: a mirror applies
    // its owner's revision, a second root on the line edits it. Either way this
    // root's manifest now reads differently, so its revision moves.
    IF _pLine^.OutImm.Revision <> _lineRevSeen THEN
        _lineRevSeen := _pLine^.OutImm.Revision;
        ConfigRev := ConfigRev + 1;
    END_IF
END_IF
_M_OeeUpdate();                                       // §8.5.1 time accounting + sampling
M_ShiftTick(Now := F_Now(), Synchronized := F_TimeSynchronized());   // §8.5.2
AlarmLog.Cyclic();                                    // §8.10 shelf auto-expiry
_M_EngineeringCyclic();                               // §7.5.2 standing gate annunciation
_healthPublisher.Cyclic(Input := _healthInput, ParCfg := _healthParCfg,
    Configured := _healthConfigured);                 // §2.7/§8.12 alarm edges + values
SystemHealth := _healthPublisher.Status;
_M_ChartRevCyclic();                                  // §3.13 coalesced chart revision
_M_HeldCyclic();                                      // §7.6.1a hold-to-run re-assert
_M_ConfigPersistCyclic();                             // §3.8b durability window
_M_DrainRestoreLoss();                                // §3.8b restore annunciation
_M_HandleHmiRequest();                                // §3.10 request mailbox
_M_DecisionCyclic();                                  // §6.11 timeout/default/overlap resolver
Access.Cyclic();
alarmActive := _M_HighestSeverity(Highest := highestSeverity);
_towerMapper.Cyclic(MachineState := MachineState, AlarmActive := alarmActive,
    HighestSeverity := highestSeverity,
    OperatorActionRequired := (Decision.Prompt <> ''),
    LampTestRequest := _lampTestRequest, ParCfg := _towerParCfg);
_lampTestRequest := FALSE;
SignalTower := _towerMapper.Status;
// §9.8 data-driven Control On/Off request endpoint. Off wins if both arrive;
// the domain/power-group implementation still validates safety, health and rearm.
ControlOnRequest := FALSE;
ControlOffRequest := FALSE;
IF ReqControlOff THEN
    ReqControlOff := FALSE;
    ReqControlOn := FALSE;
    IF Access.PermitsLogged(Gate := E_GatedAction.POWER_CONTROL) THEN
        ControlOffRequest := TRUE;
    END_IF
ELSIF ReqControlOn THEN
    ReqControlOn := FALSE;
    IF Access.PermitsLogged(Gate := E_GatedAction.POWER_CONTROL) THEN
        ControlOnRequest := TRUE;
    END_IF
END_IF
// §3.14.4 — pending mode change; §3.4.1 style decides graceful vs immediate
IF _modePend THEN
    IF _exec = E_ExecState.BUSY THEN
        IF ModePolicy[TO_INT(_mode)].Style = E_ModeSwitchStyle.GRACEFUL THEN
            _stopReq := TRUE;                             // finish the cycle at its stop point
        ELSE
            modeExitResult := OnModeExit(FirstCall := _modeExitFirst,
                RequestedMode := _modeReq);
            _modeExitFirst := FALSE;
            IF modeExitResult = 0 THEN
                OnAbort();                                // IMMEDIATE: cancel now (override may defer)
            END_IF
        END_IF
    ELSE
        IF _exec <> E_ExecState.READY THEN
            Execute := FALSE;                             // release the run command (§6.1 reset)
        ELSE
            previousMode := _mode;
            _mode := _modeReq;
            _modePend := FALSE;
            _modeExitFirst := FALSE;
            _M_CascadeMode(_mode);                        // §3.7 cascade [TC3]
            OnModeChanged(NewMode := _mode, OldMode := previousMode);
        END_IF
    END_IF
END_IF
// §8.3(c) — automatic fault capture: ERROR entry raises, ERROR exit marks gone
IF (_exec = E_ExecState.ERROR) AND (_faultEvt = 0) THEN
    _faultEvt := AlarmLog.RaiseDiag(D := _diag, ResetClass := E_ResetClass.MANUAL_RESET);
    _M_PartAborted();                  // §3.16.3: a faulted part leaves without a valid result
ELSIF (_exec <> E_ExecState.ERROR) AND (_faultEvt > 0) THEN
    AlarmLog.Gone(Slot := _faultEvt);                            // -> WAIT_RESET (blocking)
    _faultEvt := 0;
END_IF
// §6.9 — instant rollup on awaited Error; adopt a HELD child; stall as PENDING otherwise
IF _exec = E_ExecState.BUSY THEN
    IF (_awaits <> 0) AND_THEN _awaits.FaultActive THEN
        _M_FaultDiag(_awaits.GetFaultSummary());
    ELSE
        // §6.1 HELD — the held module is waiting on a condition it can name, so
        // report THAT instead of letting StallTime expire into a generic stall. A
        // declared wait is not a stall, so the watchdog stays disarmed while it lasts.
        //
        // The hold rolls up whether or not the step awaits the child (§1.1 O1: the
        // project must not have to remember a call to stay correct). `Awaits := 0`
        // says "this step owns the child's FAULT disposition" (§6.9, press AUTO
        // N200 offering scrap/return) - it does not say "stay silent while the ram
        // is HELD". A hold is recoverable information that clears itself and never
        // blocks a restart, so suppressing it only produced a Unit that sat BUSY
        // with an empty diagnostic while its own child correctly reported Held.
        // Prefer the awaited module: when a step named one it is the most specific
        // source. _M_RollupHold is called on exactly the scans the awaited branch
        // did not fire, because TwinCAT does not short-circuit and calling both
        // would let a second held child overwrite the named one.
        heldReported := FALSE;
        IF (_awaits <> 0) AND_THEN _awaits.HoldActive THEN
            _M_HoldDiag(Diag := _awaits.GetFaultSummary());
            heldReported := TRUE;
        ELSE
            heldReported := _M_RollupHold();   // §8.2 first held registered child
        END_IF
        IF heldReported THEN
            _tStall(IN := FALSE);
        ELSE
            IF Held THEN
                _M_ClearPending();     // the hold ended: drop any stall text it outlived
            END_IF
            _tStall(IN := TRUE, PT := SEL(CurrentStep.ExpectedTime > T#0S, StallTime, CurrentStep.ExpectedTime));
            IF _tStall.Q THEN
                _M_StallWalk();
            END_IF
        END_IF
    END_IF
ELSE
    _tStall(IN := FALSE);
END_IF
// §6.9(a) — every new fault joins the shift-change ring, no historian needed
_fTrig(CLK := (_exec = E_ExecState.ERROR));
_errClr(CLK := (_exec <> E_ExecState.ERROR));
IF _errClr.Q THEN
    _M_ResumeSequencesAfterError();   // §6.9 re-evaluate, do not resume blind
END_IF
IF _fTrig.Q THEN
    _M_PushHistory(_diag);
END_IF
// §8.11.4(d) — creeping WORK time is a MAINTENANCE event (Low), not downtime:
// the profiler pulses once per excursion past the configured baseline band.
IF Profiler.DegradedTrig THEN
    _M_RaiseMaintenance(Reason := E_Reason.CYCLE_TIME_DEGRADED,
        Text := 'std.maintenance.cycleTimeDegraded');
END_IF
ModeActivePublished := _mode;
RunningPublished := (_exec = E_ExecState.BUSY);
StopPendingPublished := _stopReq AND (_exec = E_ExecState.BUSY);
FOR publishIdx := 0 TO PL_Fraktal.MODE_COUNT - 1 DO
    modeIdx := publishIdx;
    SupportedModesPublished[publishIdx] := _M_Supports(Mode := modeIdx);
END_FOR
FOR publishIdx := 0 TO 2 DO
    styleIdx := publishIdx;
    SupportedRunStylesPublished[publishIdx] := _M_SupportsRunStyle(Style := styleIdx);
END_FOR
END_METHOD

// §8.13 — derive the tower input from the authoritative active-event table.
METHOD PRIVATE _M_HighestSeverity : BOOL
VAR_IN_OUT
    Highest : E_Severity;
END_VAR
VAR
    i : INT;
END_VAR
_M_HighestSeverity := FALSE;
Highest := E_Severity.LOW;
FOR i := 1 TO PL_Fraktal.MAX_ALARM_ACTIVE DO
    IF AlarmLog.Active[i].State <> E_AlarmState.CLOSED THEN
        IF NOT _M_HighestSeverity OR (AlarmLog.Active[i].Severity > Highest) THEN
            Highest := AlarmLog.Active[i].Severity;
        ELSE
            ;
        END_IF
        _M_HighestSeverity := TRUE;
    ELSE
        ;
    END_IF
END_FOR
END_METHOD

// §8.13 — remote request is MANUAL-gated and starts only while the Unit is idle.
METHOD RequestLampTest : BOOL
RequestLampTest := FALSE;
IF _exec = E_ExecState.BUSY THEN
    RETURN;
END_IF
IF NOT Access.PermitsLogged(Gate := E_GatedAction.MANUAL) THEN
    RETURN;
END_IF
_lampTestRequest := TRUE;
RequestLampTest := TRUE;
END_METHOD

// Startup station-convention seam. Runtime config writes require a registered
// typed capability; this method is not published by OPC UA.
METHOD SetSignalTowerConfig : BOOL
VAR_INPUT
    ParCfg : ST_SignalTowerParCfg;
END_VAR
IF (ParCfg.SchemaVersion <> 1) OR (ParCfg.LampTestDuration <= T#0S) THEN
    SetSignalTowerConfig := FALSE;
    RETURN;
END_IF
_towerParCfg := ParCfg;
SetSignalTowerConfig := TRUE;
END_METHOD

// TC3/platform adapter injection. Raw probe values remain OPC-UA-hidden; the
// health publisher validates and republishes the bounded status surface.
METHOD SetSystemHealth : BOOL
VAR_INPUT
    Input  : ST_SystemHealthInput;
    ParCfg : ST_SystemHealthParCfg;
END_VAR
IF ParCfg.SchemaVersion <> 1 THEN
    SetSystemHealth := FALSE;
    RETURN;
END_IF
_healthInput := Input;
_healthParCfg := ParCfg;
_healthConfigured := TRUE;
SetSystemHealth := TRUE;
END_METHOD

// §3.14 hook — one-shot after first operational scan
METHOD PROTECTED OnInit : DINT
VAR
    i : INT;
END_VAR
OnInit := SUPER^.OnInit();
_M_RestartSequences();         // §6.8 every attached chain starts at N000
SequenceViewEnabled := TRUE;   // §3.13 a Unit has a chain worth drawing;
                               // a concrete Unit may vary this per mode
Access.Setup(Provider := 0, pAlarmLog := ADR(AlarmLog)); // preserves an injected provider
_healthPublisher.Setup(SourcePath := CONCAT(Status.Name, '.SystemHealth'),
    pAlarmLog := ADR(AlarmLog));
// §3.10.2 — seed the manifest revision from boot time so every PLC restart or
// re-activation yields a NEW value (a plain counter would repeat after reboot
// and an HMI could keep a stale manifest undetected). Config writes increment.
ConfigRev := DT_TO_UDINT(F_Now());
// §3.8b — the durability provider defaults to the shipped LOCAL_RETAIN writer.
// SetConfigPersistence may already have replaced it, so this never overwrites an
// injected one.
IF _persistence = 0 THEN
    _persistence := _persistWriter;
END_IF
_liveArmed := TRUE;            // §3.8b the walk is complete: the documents may restore
// The framework's OWN station config is subject to the same rule it imposes on
// every module: version 0 is a first boot that lost nothing, any other
// unrecognized version means a real ModePolicy image was rejected and that is
// annunciated with this root's path. The base used to treat both cases as a
// silent re-initialize, which is exactly the "runs on defaults while presenting
// itself as commissioned" failure §3.8b exists to prevent.
IF NOT M_RestoreStationCfg(pVersion := ADR(_modePolicyVersion),
        SchemaVersion := MODE_POLICY_SCHEMA) THEN
    _M_InitModePolicy();
    FOR i := 0 TO PL_Fraktal.MODE_COUNT - 1 DO
        _modePolicyStored[i] := ModePolicy[i];
    END_FOR
ELSE
    FOR i := 0 TO PL_Fraktal.MODE_COUNT - 1 DO
        ModePolicy[i] := _modePolicyStored[i];
    END_FOR
END_IF
END_METHOD

// §3.14 hook — after the new mode is committed
METHOD PROTECTED OnModeChanged : DINT
VAR_INPUT
    NewMode : E_Mode;
    OldMode : E_Mode;
END_VAR
_M_HostEvent(Kind := E_HostEventKind.MODE_CHANGED, PartUid := '',
    Subject := 'Mode', Value := TO_STRING(TO_DINT(NewMode)),
    Verdict := E_Verdict.NONE, ReasonCode := E_Reason.NONE);
// §3.13 — the chart belongs to the mode that is running. A project writes nothing
// for this: it lands in the base hook every override calls SUPER^ on first (§3.14.2).
_M_ResetSequenceRows();
// §6.8 — and so do the chains: a new mode starts every chain at N000.
_M_RestartSequences();
OnModeChanged := 0;
END_METHOD

// Core §11.6: CHANGEOVER starts when its guided sequence actually starts, not
// merely when the operator selects the mode or transactionally loads a model.
METHOD PROTECTED OnCommandStart : DINT
OnCommandStart := SUPER^.OnCommandStart();
IF _mode = E_Mode.CHANGEOVER THEN
    _M_HostEvent(Kind := E_HostEventKind.CHANGEOVER_STARTED, PartUid := '',
        Subject := 'Model', Value := Model.ModelCode,
        Verdict := E_Verdict.NONE, ReasonCode := E_Reason.NONE);
END_IF
END_METHOD

// §3.14.4 — called every scan while a mode request is pending and the Unit is BUSY.
// Return 0 = consent to immediate cancel (default); >0 = still stopping gracefully.
METHOD PROTECTED OnModeExit : DINT
VAR_INPUT
    FirstCall : BOOL;
    RequestedMode : E_Mode;
END_VAR
OnModeExit := 0;
END_METHOD

// §8.3(b) — deliberate operator reset of blocking events (release-gated per §7.6/§14).
// ONE operator action has to make the Unit restartable, so this closes the blocking
// events AND clears the latched control state they were reporting: see _M_RecoverState.
METHOD OperatorReset : BOOL
IF NOT Access.PermitsLogged(Gate := E_GatedAction.ALARM_RESET) THEN
    OperatorReset := FALSE;            // §7.7
    RETURN;
END_IF
OperatorReset := _M_RecoverState();
OperatorReset := AlarmLog.OperatorReset() OR OperatorReset;
END_METHOD

// §8.3(b)/§6.1 — the control-state half of a reset. Closing the alarm alone left the
// machine locked: the Unit's run command and the child commands its mode chain had
// issued both stayed asserted, and §6.1's Execute-drop reset — the only exit from a
// latched terminal state — needs them LOW. A frozen chain cannot drop them itself,
// because a Unit that is not BUSY never calls _M_Dispatch again, so the step holding
// `child.Execute := TRUE` never runs. Nothing else in the system clears it, and the
// next Start re-issues the same already-TRUE input: no rising edge, the child stays
// in ERROR, and the Unit re-adopts the fault through the §8.2 rollup. That is the
// press hard-lock. Returns TRUE when there was something to recover.
// Deliberately does NOT clear ERROR here: Cyclic keeps that ownership (§6.1), so a
// cause that is still live re-faults on the next command edge instead of vanishing.
METHOD PROTECTED _M_RecoverState : BOOL
_M_RecoverState := FALSE;
IF (_exec <> E_ExecState.ERROR) AND NOT AlarmLog.Blocking THEN
    RETURN;                            // nothing latched: a stray reset changes nothing
END_IF
OnOperatorReset();                     // §3.14 hook: withdraw outputs, reset mode chains
_M_ReleaseChildCommands();             // stranded child commands -> READY next scan
_M_ClearPending();
_stopReq := FALSE;
IF _exec = E_ExecState.BUSY THEN
    // Defined safe reaction (§5.6) for a blocking event raised by application code
    // while the mode chain still runs: a recovery reset cancels what was running
    // rather than leaving a chain we just reset still driving the machine.
    AbortCommand();
END_IF
Execute  := FALSE;                     // stale run command -> Unit READY next scan
_faultEvt := 0;                        // the event is closed here, not by a later Gone()
_M_RecoverState := TRUE;
END_METHOD

// §3.14 hook — an accepted operator reset is recovering this Unit. Override to
// withdraw application outputs and reset application-owned mode chains before the
// base releases the run command; call SUPER^.OnOperatorReset() first (§3.14.2).
// Called only when something was actually latched (ERROR or a blocking alarm), so an
// override may assume it is a recovery, not a routine poll.
METHOD PROTECTED OnOperatorReset : DINT
OnOperatorReset := 0;
END_METHOD

// Application-only seam for an ordinary hardwired fault-reset/acknowledge button,
// mirroring RequestLocalControl (§9.8): it is a METHOD, not OPC UA data, so remote
// clients still go through the access-gated OPERATOR_RESET request and cannot reach
// this path. A cabinet button IS its own authorization (physical presence), so it
// carries no §7.7 session check — but the reset is still audited as a §8.3 event,
// and it recovers exactly the same state as an operator reset, never more.
// The composition root calls this from its hardware driver on the button's rising
// edge, once per root Unit it should clear.
METHOD RequestLocalReset : BOOL
VAR
    auditSlot : INT;
END_VAR
auditSlot := AlarmLog.Raise(Reason := E_Reason.NONE,
    Text := 'std.audit.localResetRequested', Source := _name,
    Severity := E_Severity.LOW, Category := E_Category.SYSTEM,
    ResetClass := E_ResetClass.AUTO_RESET);
IF auditSlot > 0 THEN AlarmLog.Gone(Slot := auditSlot); END_IF
RequestLocalReset := _M_RecoverState();
RequestLocalReset := AlarmLog.OperatorReset() OR RequestLocalReset;
END_METHOD

// §3.8 optional HMI/MES selection catalog. Recipe providers remain pluggable;
// the application registers only the model identities it deliberately exposes.
METHOD RegisterAvailableModel : BOOL
VAR_INPUT
    Id : ST_ModelId;
END_VAR
VAR
    i : INT;
END_VAR
RegisterAvailableModel := FALSE;
IF (Id.ModelCode = '') OR (AvailableModelCount >= PL_Fraktal.MAX_RECIPES) THEN
    RETURN;
END_IF
FOR i := 1 TO AvailableModelCount DO
    IF AvailableModels[i].ModelCode = Id.ModelCode THEN
        RETURN;
    END_IF
END_FOR
AvailableModels[AvailableModelCount + 1] := Id;
AvailableModelCount := AvailableModelCount + 1;
ConfigRev := ConfigRev + 1;    // §3.10.2 — manifest changed
RegisterAvailableModel := TRUE;
END_METHOD

// §9.8 remote control-domain request. The acknowledgement is the result of this
// authorization check; it is never reported accepted before POWER_CONTROL runs.
METHOD RequestControlPower : BOOL
VAR_INPUT
    ControlOn : BOOL;
END_VAR
RequestControlPower := FALSE;
IF NOT Access.PermitsLogged(Gate := E_GatedAction.POWER_CONTROL) THEN
    RETURN;
END_IF
IF ControlOn THEN
    ReqControlOn := TRUE;
    ReqControlOff := FALSE;
ELSE
    ReqControlOff := TRUE;                         // Off wins if both were requested
    ReqControlOn := FALSE;
END_IF
RequestControlPower := TRUE;
END_METHOD

// §6.11 authoritative decision entry. START_STOP is the access gate because the
// answer advances a running Unit chain; option-specific process releases append
// through _M_AppendDecisionInterlocks. A stale/invalid answer never latches.
METHOD SubmitDecision : BOOL
VAR_INPUT
    Option : INT;
END_VAR
VAR_IN_OUT
    Report : ST_ReleaseReport;
END_VAR
Report.Count := 0;
Report.Released := FALSE;
SubmitDecision := FALSE;
IF NOT Access.PermitsLogged(Gate := E_GatedAction.START_STOP) THEN
    _M_AddReason(Report := Report, Text := 'std.release.insufficientStartStop',
        Reason := E_Reason.NONE, Kind := E_ReleaseKind.ACCESS);
END_IF
IF (_exec <> E_ExecState.BUSY) OR (Decision.Prompt = '') THEN
    _M_AddReason(Report := Report, Text := 'std.release.noActiveDecision',
        Reason := E_Reason.NONE, Kind := E_ReleaseKind.OTHER);
ELSIF (Option < 1) OR (Option > PL_Fraktal.MAX_OPTIONS) THEN
    _M_AddReason(Report := Report, Text := 'std.release.invalidDecisionOption',
        Reason := E_Reason.UNSUPPORTED_COMMAND, Kind := E_ReleaseKind.OTHER);
ELSIF Decision.Options[Option] = '' THEN
    _M_AddReason(Report := Report, Text := 'std.release.invalidDecisionOption',
        Reason := E_Reason.UNSUPPORTED_COMMAND, Kind := E_ReleaseKind.OTHER);
ELSE
    _M_AppendDecisionInterlocks(Option := Option, Report := Report);
END_IF
Report.Released := (Report.Count = 0);
IF Report.Released THEN
    DecisionAnswer := Option;
    SubmitDecision := TRUE;
END_IF
END_METHOD

// §7.7 persistent per-root policy edit. The policy's own ACCESS_POLICY threshold
// is rechecked before any threshold — including itself — can change.
METHOD SetAccessLevel : BOOL
VAR_INPUT
    Gate : E_GatedAction;
    Level : E_AccessLevel;
END_VAR
SetAccessLevel := FALSE;
IF NOT Access.PermitsLogged(Gate := E_GatedAction.ACCESS_POLICY) THEN
    RETURN;
END_IF
// Never allow an anonymous/lower session to raise the policy above itself and
// strand the retained station configuration without a usable administrator.
IF (Gate = E_GatedAction.ACCESS_POLICY) AND (Level > Access.CurrentLevel) THEN
    RETURN;
END_IF
SetAccessLevel := Access.ConfigureRequired(Gate := Gate, Level := Level);
IF SetAccessLevel THEN
    ConfigRev := ConfigRev + 1;
END_IF
END_METHOD

// §7.7 persistent idle timeout (0 = never), self-gated by ACCESS_POLICY.
METHOD SetSessionTimeout : BOOL
VAR_INPUT
    TimeoutMs : UDINT;
END_VAR
SetSessionTimeout := FALSE;
IF NOT Access.PermitsLogged(Gate := E_GatedAction.ACCESS_POLICY) THEN
    RETURN;
END_IF
SetSessionTimeout := Access.ConfigureSessionTimeout(TimeoutMs := TimeoutMs);
IF SetSessionTimeout THEN
    ConfigRev := ConfigRev + 1;
END_IF
END_METHOD

// §3.8a/§7.7 centralized HMI configuration authority. Concrete overrides never
// need to remember DATA_WRITE or root ownership; they validate only their field.
METHOD WriteConfig : BOOL
VAR_INPUT
    TargetPath : STRING(255);
    WriteKey : STRING(160);
    Revision : DINT;
    TextValue : STRING(255);
END_VAR
WriteConfig := FALSE;
IF NOT _M_ConfigRestored() THEN
    RETURN;                            // §3.8b the restore would replay over it
END_IF
IF (WriteKey = '') OR (Revision <= 0)
OR NOT _M_OwnsModulePath(Path := TargetPath) THEN
    RETURN;
END_IF
// §3.8d - the VALUE's effective write level (its class, raised by its own
// minimum); DATA_WRITE for a value in the built-in class, as before.
IF NOT Access.M_PermitsLevelLogged(Required := _M_DataLevelOf(TargetPath := TargetPath,
        WriteKey := WriteKey, ForWrite := TRUE)) THEN
    RETURN;
END_IF
WriteConfig := _M_WriteBaseConfig(TargetPath := TargetPath, WriteKey := WriteKey,
    Revision := TO_UDINT(Revision), TextValue := TextValue, Commit := TRUE);
IF NOT WriteConfig THEN
    WriteConfig := _M_RouteConfigWrite(TargetPath := TargetPath,
        WriteKey := WriteKey, Revision := TO_UDINT(Revision), TextValue := TextValue);
END_IF
// §3.8a - a model-data value lives in a recipe record too. Another model's edit
// exists ONLY in that record, so failing to save it fails the write; the active
// model's edit is already live, and saving it keeps it across a changeover.
IF WriteConfig AND (TargetPath = Status.Name) AND _M_ModelScopedKey(WriteKey := WriteKey) THEN
    IF NOT _M_SaveModelData() AND (_pModelView <> 0) THEN
        WriteConfig := FALSE;
    END_IF
END_IF
IF WriteConfig THEN
    ConfigRev := ConfigRev + 1;
    _M_MarkPersistPending();           // §3.8b: accepted is LIVE, not yet DURABLE
END_IF
END_METHOD

// §3.8c - the root authority for a capture. Deliberately the same gate, the same
// ownership check and the same ConfigRev bump as WriteConfig: a capture is a
// write whose value came from the machine, and it is no more and no less
// privileged than one the operator typed (§3.8c(d)).
METHOD CaptureConfig : BOOL
VAR_INPUT
    TargetPath : STRING(255);
    WriteKey   : STRING(160);
    Revision   : DINT;
END_VAR
CaptureConfig := FALSE;
IF NOT _M_ConfigRestored() THEN
    RETURN;
END_IF
IF (WriteKey = '') OR (Revision <= 0)
OR NOT _M_OwnsModulePath(Path := TargetPath) THEN
    RETURN;
END_IF
IF NOT Access.M_PermitsLevelLogged(Required := _M_DataLevelOf(TargetPath := TargetPath,
        WriteKey := WriteKey, ForWrite := TRUE)) THEN
    RETURN;
END_IF
// Framework-owned keys offer no capture: they are policy, not measurements.
CaptureConfig := M_ApplyCapture(Scope := TargetPath, WriteKey := WriteKey,
    Revision := TO_UDINT(Revision), RootReady := (_exec = E_ExecState.READY));
IF CaptureConfig THEN
    ConfigRev := ConfigRev + 1;
END_IF
END_METHOD

// Core §7.5.1 — inject the station's commissioning/engineering gate register at
// Setup, the same shape as SetPartCarrier. Wiring it is what makes the §7.5.2
// standing annunciation appear and what arms the §10.5.1 force surface; a Unit
// with no register is a production Unit and both are simply absent.
//
// Declaring the framework's OWN force gate happens here rather than in the
// project, so a composition root that wires the register cannot forget it
// (§1.1 O1) and cannot arm forcing without also annunciating it.
METHOD SetEngineeringMode
VAR_INPUT
    Mode : REFERENCE TO FB_EngineeringMode;
END_VAR
_engineering REF= Mode;
IF __ISVALIDREF(_engineering) THEN
    _engineering.M_DeclareOutputForcing();
ELSE
    ;
END_IF
END_METHOD

// Core §10.5.1 rules 1 and 3 — may a held force set-point be applied to this
// Unit's outputs right now? The project hardware driver passes the result to
// FB_IoTopologyPublisher.M_ApplyForces every scan, and ForceChannel gates the
// operator request on the identical predicate, so "accepted" and "applied" can
// never disagree. Everything else about a force (access, ownership, direction,
// mapping) is proved elsewhere; this is only the build gate and the mode/state.
METHOD M_ForcePermitted : BOOL
M_ForcePermitted := FALSE;
IF NOT __ISVALIDREF(_engineering) THEN
    RETURN;
END_IF
IF NOT _engineering.ForcingActive THEN
    RETURN;
END_IF
// A running module reasserts its own outputs, so a force is only honest while
// the Unit is idle in MANUAL; leaving either withdraws every force (§10.5.1(3)).
M_ForcePermitted := (_mode = E_Mode.MANUAL) AND (_exec = E_ExecState.READY);
END_METHOD

// Core §7.5.2 — the standing annunciation: one LOW/SYSTEM/AUTO_RESET event per
// registered gate, for as long as that gate is registered.
//
// Why each choice is the way it is, because every one of them is load-bearing:
//   AUTO_RESET  a MANUAL_RESET event refuses Start (§8.3(b)), which would make
//               commissioning gates block the commissioning they exist to serve;
//   LOW/SYSTEM  the lowest priority and the lowest risk class - this says how the
//               software was BUILT, not that the process or safety is impaired,
//               and a louder class would displace real alarms (§8.9);
//   unclearable OperatorReset only closes MANUAL_RESET events, so no operator
//               action reaches this one, and its §8.9 record is not shelvable, so
//               §8.10 cannot silence it either. It closes when the gate is gone -
//               which, gates being build constants, means a new download.
METHOD PRIVATE _M_EngineeringCyclic
VAR
    i : INT;
    gateCount : INT;
END_VAR
IF NOT __ISVALIDREF(_engineering) THEN
    RETURN;
END_IF
gateCount := _engineering.Count;
IF gateCount > PL_Fraktal.MAX_ENGINEERING_GATES THEN
    gateCount := PL_Fraktal.MAX_ENGINEERING_GATES;
END_IF
FOR i := 1 TO gateCount DO
    // Self-healing on purpose. If this slot were ever closed and reused by
    // another event, a remembered index would leave the annunciation silently
    // absent for the rest of the run - the one failure mode a non-clearable
    // message must not have. Re-verify identity, then re-raise.
    IF _engineeringEvt[i] > 0 THEN
        IF (AlarmLog.Active[_engineeringEvt[i]].State = E_AlarmState.CLOSED)
        OR (AlarmLog.Active[_engineeringEvt[i]].ReasonCode <> E_Reason.COMMISSIONING_GATE_ACTIVE) THEN
            _engineeringEvt[i] := 0;
        ELSE
            ;
        END_IF
    ELSE
        ;
    END_IF
    IF _engineeringEvt[i] = 0 THEN
        _engineeringEvt[i] := AlarmLog.Raise(Reason := E_Reason.COMMISSIONING_GATE_ACTIVE,
            Text := _engineering.Gates[i].DescriptionKey, Source := _name,
            Severity := E_Severity.LOW, Category := E_Category.SYSTEM,
            ResetClass := E_ResetClass.AUTO_RESET);
    ELSE
        ;
    END_IF
END_FOR
END_METHOD

// §10.5.1 centralized force authority. Only an idle MANUAL Unit may reach the
// application resolver; that resolver still proves root ownership, OUTPUT,
// non-safety identity, mapping and the channel-specific release.
METHOD ForceChannel : BOOL
VAR_INPUT
    ChannelPath : STRING(255);
    Force : BOOL;
    BoolText : STRING(255);
    AnalogText : STRING(160);
END_VAR
ForceChannel := FALSE;
IF NOT Access.PermitsLogged(Gate := E_GatedAction.MANUAL) THEN
    RETURN;
END_IF
// §10.5.1 rules 1 and 3 in one predicate, the same one the hardware driver
// applies each scan - so the request can never be accepted under conditions
// under which the force would not actually be applied.
IF NOT M_ForcePermitted() OR (ChannelPath = '') THEN
    RETURN;
END_IF
ForceChannel := _M_RouteForceChannel(ChannelPath := ChannelPath, Force := Force,
    BoolText := BoolText, AnalogText := AnalogText);
END_METHOD

// Core §7.8 — full rollup for the simpler gated Unit actions (Stop, ALARM_RESET,
// CHANGEOVER, MODE_CHANGE, step). Same predicate the gates use. Start has its own
// richer ReleaseReportStart (interlocks); manual has ReleaseReportManual (target).
METHOD ReleaseReportAction : BOOL
VAR_INPUT
    Gate : E_GatedAction;
END_VAR
VAR_IN_OUT
    Report : ST_ReleaseReport;
END_VAR
Report.Count := 0;
Report.Released := FALSE;
// access is the common gate
IF NOT Access.Permits(Gate := Gate) THEN
    _M_AddReason(Report := Report, Text := 'std.release.insufficientAction', Reason := E_Reason.NONE, Kind := E_ReleaseKind.ACCESS);
END_IF
// per-action state preconditions
CASE Gate OF
    E_GatedAction.CHANGEOVER:
        IF _exec = E_ExecState.BUSY THEN
            _M_AddReason(Report := Report, Text := 'std.release.changeoverRunning', Reason := E_Reason.NONE, Kind := E_ReleaseKind.MODE);
        END_IF
    E_GatedAction.ALARM_RESET:
        IF NOT AlarmLog.Blocking THEN
            _M_AddReason(Report := Report, Text := 'std.release.noBlockingAlarm', Reason := E_Reason.NONE, Kind := E_ReleaseKind.OTHER);
        END_IF
    E_GatedAction.MODE_CHANGE:
        IF _modePend THEN
            _M_AddReason(Report := Report, Text := 'std.release.modeChangeAlreadyPending', Reason := E_Reason.NONE, Kind := E_ReleaseKind.MODE);
        ELSIF (_exec = E_ExecState.BUSY)
        AND (ModePolicy[TO_INT(_mode)].Shield = E_ModeSwitchShield.BLOCKED_WHILE_RUNNING) THEN
            _M_AddReason(Report := Report, Text := 'std.release.modeSwitchBlockedWhileRunning',
                Reason := E_Reason.NONE, Kind := E_ReleaseKind.MODE);
        ELSE
            ;
        END_IF
ELSE
    ;                                          // actions with no extra state predicate
END_CASE
Report.Released := (Report.Count = 0);
ReleaseReportAction := Report.Released;
END_METHOD

// Core §7.8 — full rollup of why a manual command to Target would be refused (§7.6.1).
METHOD ReleaseReportManual : BOOL
VAR_INPUT
    TargetPath : STRING(255);
    Value : DINT;
END_VAR
VAR_IN_OUT
    Report : ST_ReleaseReport;
END_VAR
Report.Count := 0;
Report.Released := FALSE;
IF _mode <> E_Mode.MANUAL THEN
    _M_AddReason(Report := Report, Text := 'std.release.manualModeRequired', Reason := E_Reason.NONE, Kind := E_ReleaseKind.MODE);
END_IF
IF NOT Access.Permits(Gate := E_GatedAction.MANUAL) THEN
    _M_AddReason(Report := Report, Text := 'std.release.insufficientManual', Reason := E_Reason.NONE, Kind := E_ReleaseKind.ACCESS);
END_IF
_M_AppendManualInterlocks(TargetPath := TargetPath, Value := Value, Report := Report);  // §7.6, target+command-aware
Report.Released := (Report.Count = 0);
ReleaseReportManual := Report.Released;
END_METHOD

// Core §7.8 — pure query: the FULL rollup of why Start would be refused right now.
// This is the authoritative machine predicate consumed by Start (no drift).
// Released = TRUE means Start proceeds. Lists mode + access + blocking-alarm,
// control-domain, and concrete mode-entry release reasons. The caller owns the
// bounded report storage; returning this large record by value can overflow a
// TwinCAT task stack when Start consumes the result.
METHOD ReleaseReportStart : BOOL
VAR_IN_OUT
    Report : ST_ReleaseReport;
END_VAR
Report.Count := 0;
Report.Released := FALSE;
// access (§7.7)
IF NOT Access.Permits(Gate := E_GatedAction.START_STOP) THEN
    _M_AddReason(Report := Report, Text := 'std.release.insufficientStartStop', Reason := E_Reason.NONE, Kind := E_ReleaseKind.ACCESS);
END_IF
// mode / run state (§3.4)
IF _modePend THEN
    _M_AddReason(Report := Report, Text := 'std.release.modeChangePending', Reason := E_Reason.NONE, Kind := E_ReleaseKind.MODE);
END_IF
IF _mode = E_Mode.MANUAL THEN
    _M_AddReason(Report := Report, Text := 'std.release.manualHasNoAutoSequence', Reason := E_Reason.NONE, Kind := E_ReleaseKind.MODE);
END_IF
IF _exec <> E_ExecState.READY THEN
    _M_AddReason(Report := Report, Text := 'std.release.unitNotReady', Reason := E_Reason.NONE, Kind := E_ReleaseKind.MODE);
END_IF
// blocking alarm (§8.3)
IF AlarmLog.Blocking THEN
    _M_AddReason(Report := Report, Text := 'std.release.manualReset', Reason := E_Reason.NONE, Kind := E_ReleaseKind.ALARM);
END_IF
// lost configuration image (§3.8b): the DEPLOYMENT's declared consequence. The
// policy was stored and published but read nowhere, so a station that declared
// BLOCK_UNTIL_ACKNOWLEDGED started on defaults anyway. This is where it is read.
IF ConfigPersist.RestoreLost AND NOT ConfigPersist.RestoreAcknowledged
AND (ConfigPersist.RestorePolicy = E_ConfigRestorePolicy.BLOCK_UNTIL_ACKNOWLEDGED) THEN
    _M_AddReason(Report := Report, Text := 'std.release.configRestoreUnacknowledged', Reason := E_Reason.CONFIG_RESTORE_LOST, Kind := E_ReleaseKind.ALARM);
END_IF
// §3.8b - the live documents are still being read back: the running values are
// not yet the ones last made durable.
IF NOT _M_ConfigRestored() THEN
    _M_AddReason(Report := Report, Text := 'std.release.configRestoring', Reason := E_Reason.NONE, Kind := E_ReleaseKind.OTHER);
END_IF
IF ControlDomain.Present AND NOT ControlDomain.ReadyForStart THEN
    _M_AddReason(Report := Report, Text := 'std.release.controlDomainNotReady', Reason := E_Reason.NONE, Kind := E_ReleaseKind.INTERLOCK);
END_IF
// active mode's immediate entry/frontier conditions (concrete override)
_M_AppendInterlocks(Report := Report);
Report.Released := (Report.Count = 0);
ReleaseReportStart := Report.Released;
END_METHOD

// §8.5.1 — clear accumulators + ring (shift start). Gated: §7.7 DATA_WRITE; audited §8.3.
METHOD ResetOee : BOOL
VAR
    i : INT;
    auditSlot : INT;
END_VAR
IF NOT Access.PermitsLogged(Gate := E_GatedAction.DATA_WRITE) THEN
    ResetOee := FALSE;
    RETURN;
END_IF
_oeeGoodBase := GoodCount;
_oeeNokBase := NokCount;
Oee.RunMs := 0; Oee.DownMs := 0; Oee.IdleMs := 0;
FOR i := 1 TO PL_Fraktal.MAX_OEE_SAMPLES DO
    OeeTrend[i].Oee := 0.0; OeeTrend[i].OeeValid := FALSE;
    OeeTrend[i].Availability := 0.0; OeeTrend[i].Performance := 0.0; OeeTrend[i].Quality := 0.0;
END_FOR
OeeTrendHead := 0;
_oeeSampMs := 0;
_M_OeeCompute();
_shiftManualReset := TRUE;                  // §8.5.2(c): the shift record will say so
auditSlot := AlarmLog.Raise(Reason := E_Reason.NONE,
    Text := 'std.audit.oeeReset', Source := _name,
    Severity := E_Severity.LOW, Category := E_Category.SYSTEM, ResetClass := E_ResetClass.AUTO_RESET);
IF auditSlot > 0 THEN AlarmLog.Gone(Slot := auditSlot); END_IF
ResetOee := TRUE;
END_METHOD

// §3.4.2 — HMI HOLD_TO_RUN input. NON-SAFETY (§9): never a dead-man; interlocks
// still apply at every step. TRUE only while the operator holds the button.
METHOD SetHoldRun : BOOL
VAR_INPUT
    Held : BOOL;
END_VAR
IF Held AND (NOT Access.PermitsLogged(Gate := E_GatedAction.START_STOP)
OR (RunStyle <> E_RunStyle.HOLD_TO_RUN) OR (_exec <> E_ExecState.BUSY)) THEN
    SetHoldRun := FALSE;
    RETURN;
END_IF
_holdRun := Held;                     // FALSE is always accepted so a hold cannot stick
SetHoldRun := TRUE;
END_METHOD

// §8.5.1 — configure the ideal cycle time (per model, §3.8). 0 disables Performance.
METHOD SetIdealCycle : BOOL
VAR_INPUT
    Ms : UDINT;
END_VAR
Oee.IdealCycleMs := Ms;
SetIdealCycle := TRUE;
END_METHOD

// §3.4/§3.7 — FALSE = unsupported (graceful rejection); TRUE = committed or pending
METHOD SetMode : BOOL
VAR_INPUT
    Mode : E_Mode;
END_VAR
IF NOT Access.PermitsLogged(Gate := E_GatedAction.MODE_CHANGE) THEN
    SetMode := FALSE;                  // §7.7(c): who-gate ANDs the machine gates
    RETURN;
END_IF
IF NOT _M_Supports(Mode) THEN
    SetMode := FALSE;
    RETURN;
END_IF
IF (Mode = _mode) AND NOT _modePend THEN
    SetMode := TRUE;
    RETURN;
END_IF
// §3.4.1 shield: policy of the mode being LEFT governs while its sequence runs
IF (_exec = E_ExecState.BUSY)
AND (ModePolicy[TO_INT(_mode)].Shield = E_ModeSwitchShield.BLOCKED_WHILE_RUNNING) THEN
    SetMode := FALSE;                  // must Stop first (graceful rejection, not a fault)
    RETURN;
END_IF
IF (NOT _modePend) OR (_modeReq <> Mode) THEN
    _modeExitFirst := TRUE;
END_IF
_modeReq := Mode;
_modePend := TRUE;
SetMode := TRUE;
END_METHOD

// §3.1b/§3.8 — transactional model change: prepare the whole subtree, then commit.
METHOD SetModel : BOOL
VAR_INPUT
    Id : ST_ModelId;
END_VAR
IF NOT Access.PermitsLogged(Gate := E_GatedAction.CHANGEOVER) THEN
    SetModel := FALSE;                 // §7.7
    RETURN;
END_IF
IF _exec = E_ExecState.BUSY THEN
    SetModel := FALSE;                 // changeover is not mid-cycle (§3.8 loads at CHANGEOVER)
    RETURN;
END_IF
IF NOT PrepareRecipe(Model := Id) THEN
    AbortRecipe();
    SetModel := FALSE;
    RETURN;
END_IF
CommitRecipe();                         // infallible after successful preparation
Model := Id;                           // identity changes only after subtree commit
ConfigRev := ConfigRev + 1;            // §3.10.2 — recipe/config leaves changed
SetModel := TRUE;
END_METHOD

// §11.6.1 internal composition seam; not a remote command surface.
METHOD M_PublishMaterialChanged : BOOL
VAR_INPUT
    Material : STRING(80);
    Value    : STRING(80);
END_VAR
M_PublishMaterialChanged := _M_HostEvent(
    Kind := E_HostEventKind.MATERIAL_CHANGED, PartUid := '', Subject := Material,
    Value := Value, Verdict := E_Verdict.NONE, ReasonCode := E_Reason.NONE);
END_METHOD

// §11.6.1 internal composition seam; not a remote command surface.
METHOD M_PublishToolChanged : BOOL
VAR_INPUT
    Tool  : STRING(80);
    Value : STRING(80);
END_VAR
M_PublishToolChanged := _M_HostEvent(
    Kind := E_HostEventKind.TOOL_CHANGED, PartUid := '', Subject := Tool,
    Value := Value, Verdict := E_Verdict.NONE, ReasonCode := E_Reason.NONE);
END_METHOD

// §11.6.2 inject an optional OPC UA/MES/REST/MQTT delivery adapter.
METHOD M_SetHostEventSink : BOOL
VAR_INPUT
    Sink : I_HostEventSink;
END_VAR
M_SetHostEventSink := HostEvents.SetSink(Sink := Sink);
END_METHOD

// §3.16.2 — inject the part carrier at the composition root (0 = traceability off).
// Source-agnostic: BY_POSITION local, RFID, DataMatrix, or host, behind I_PartCarrier.
METHOD SetPartCarrier : BOOL
VAR_INPUT
    Carrier : I_PartCarrier;
END_VAR
_carrier := Carrier;
SetPartCarrier := (Carrier <> 0);
END_METHOD

// §3.4.2 — HMI selects the run style for the active mode. Modes that don't opt in
// (see _M_SupportsRunStyle) reject non-CONTINUOUS. Access: MODE_CHANGE-gated (§7.7).
METHOD SetRunStyle : BOOL
VAR_INPUT
    Style : E_RunStyle;
END_VAR
IF NOT Access.PermitsLogged(Gate := E_GatedAction.MODE_CHANGE) THEN
    SetRunStyle := FALSE;
    RETURN;
END_IF
IF (Style <> E_RunStyle.CONTINUOUS) AND NOT _M_SupportsRunStyle(Style := Style) THEN
    SetRunStyle := FALSE;               // mode didn't opt into stepping (graceful reject)
    RETURN;
END_IF
RunStyle := Style;
SetRunStyle := TRUE;
END_METHOD

// §8.10 — gated HMI entry: shelve an active alarm's ANNUNCIATION (control untouched).
// §7.7 ALARM_SHELVE + audit; refuses SAFETY / unrationalized reasons (AlarmLog rules).
METHOD ShelveAlarm : BOOL
VAR_INPUT
    Slot      : INT;
    DurationS : UDINT;
END_VAR
IF NOT Access.PermitsLogged(Gate := E_GatedAction.ALARM_SHELVE) THEN
    ShelveAlarm := FALSE;
    RETURN;
END_IF
ShelveAlarm := AlarmLog.Shelve(Slot := Slot, DurationS := DurationS);
END_METHOD

// §3.3/§6 intro — the run IS a §6.1 command.
// §7.8: ReleaseReportStart is the authoritative machine gate as well as the
// operator explanation, so a concrete Unit cannot report an interlock it ignores.
// Build directly into the published response storage: ST_ReleaseReport is too
// large for nested by-value/local copies on a small TwinCAT task stack.
METHOD Start : BOOL
IF NOT Access.PermitsLogged(Gate := E_GatedAction.START_STOP) THEN
    Start := FALSE;                    // §7.7
    RETURN;
END_IF
IF ReleaseReportStart(Report := HmiResponse.Report) THEN
    _stopReq := FALSE;                 // §8.3(b): a MANUAL_RESET event blocks restart
    Execute := TRUE;
    Start := TRUE;
ELSE
    Start := FALSE;
END_IF
END_METHOD

// §3.4.2 — HMI single-step: request advance of one step (edge-consumed by _M_StepGate).
METHOD StepRequest : BOOL
IF NOT Access.PermitsLogged(Gate := E_GatedAction.START_STOP)
OR (RunStyle <> E_RunStyle.SINGLE_STEP) OR (_exec <> E_ExecState.BUSY) THEN
    StepRequest := FALSE;
    RETURN;
END_IF
_stepReq := TRUE;
StepRequest := TRUE;
END_METHOD

// §3.3 — stop after the current cycle
METHOD Stop : BOOL
IF NOT Access.PermitsLogged(Gate := E_GatedAction.START_STOP) THEN
    Stop := FALSE;                     // §7.7
    RETURN;
END_IF
IF _exec = E_ExecState.BUSY THEN
    _stopReq := TRUE;
ELSE
    _stopReq := FALSE;
    Execute := FALSE;                  // release a terminal run command (ERROR/DONE/ABORTED)
END_IF
Stop := TRUE;
END_METHOD

// §3.4 — TRUE while a stop is requested but the sequence is still finishing
// (running -> stopping). HMI blinks the stop button on this.
PROPERTY StopPending : BOOL
GET
StopPending := _stopReq AND (_exec = E_ExecState.BUSY);
END_GET
END_PROPERTY

// §8.10 — gated HMI entry: restore annunciation.
METHOD UnshelveAlarm : BOOL
VAR_INPUT
    Slot : INT;
END_VAR
IF NOT Access.PermitsLogged(Gate := E_GatedAction.ALARM_SHELVE) THEN
    UnshelveAlarm := FALSE;
    RETURN;
END_IF
UnshelveAlarm := AlarmLog.Unshelve(Slot := Slot);
END_METHOD

METHOD PRIVATE _M_SyncModelCatalog
VAR
    i : INT;
    j : INT;
    id : ST_ModelId;
    exists : BOOL;
    found : UINT;
    info : ST_ConfigSetInfo;
    record : ST_ConfigRecord;
END_VAR
IF _modelCatalog = 0 THEN ModelCapacity := 0; RETURN; END_IF
IF _modelCatalogSeen = _modelCatalog.M_ModelCount(RecipeKey := _modelKey) THEN RETURN; END_IF
_modelCatalogSeen := _modelCatalog.M_ModelCount(RecipeKey := _modelKey);
FOR i := 1 TO _modelCatalog.M_ModelCount(RecipeKey := _modelKey) DO
    IF _modelCatalog.M_ModelAt(RecipeKey := _modelKey, Index := i, Id := id) THEN
        exists := FALSE;
        FOR j := 1 TO AvailableModelCount DO
            IF AvailableModels[j].ModelCode = id.ModelCode THEN exists := TRUE; END_IF
        END_FOR
        IF NOT exists THEN RegisterAvailableModel(Id := id); END_IF
    END_IF
END_FOR
ModelCapacity := _modelCatalog.M_ModelCapacity(RecipeKey := _modelKey);
IF ModelCapacity > PL_Fraktal.MAX_RECIPES THEN ModelCapacity := PL_Fraktal.MAX_RECIPES; END_IF
IF _modelCatalog.M_TakeCatalogRestoreLoss(Found => found) THEN
    _restoreLost := TRUE;
    _restoreFound := found;
    _restoreExpected := 1;
END_IF
IF NOT _M_CaptureConfig(SetName := '_validation', Kind := E_ConfigKind.PAR_CFG, ModelIndex := 0) THEN
    ModelCapacity := 0; RETURN;
END_IF
_snapshot.M_ReadInfo(SetName := '_validation', Info := info);
FOR i := 1 TO info.RecordCount DO
    _snapshot.M_ReadRecord(SetName := '_validation', Index := i, Record := record);
    IF NOT _M_OwnsModelRecord(Record := record) THEN ModelCapacity := 0; EXIT; END_IF
END_FOR
END_METHOD

METHOD PRIVATE _M_OwnsModelRecord : BOOL
VAR_INPUT
    Record : ST_ConfigRecord;
END_VAR
VAR
    i : INT;
END_VAR
_M_OwnsModelRecord := FALSE;
IF (Record.Scope <> Status.Name) OR (Record.Kind <> E_ConfigKind.PAR_CFG) THEN RETURN; END_IF
FOR i := 1 TO _nConfigWrite DO
    IF _pConfigWrite[i - 1].Key = Record.WriteKey THEN
        _M_OwnsModelRecord := (_pConfigWrite[i - 1].Kind = E_ConfigKind.PAR_CFG)
            AND (_pConfigWrite[i - 1].pTarget >= _pModelRegion)
            AND (_pConfigWrite[i - 1].pTarget < _pModelRegion + _modelRegionSize);
        RETURN;
    END_IF
END_FOR
END_METHOD

// Freeze untrusted storage before validation or a commit pass.
METHOD PRIVATE _M_CopySet : BOOL
VAR_INPUT
    SetName : STRING(80);
END_VAR
VAR
    info : ST_ConfigSetInfo;
    record : ST_ConfigRecord;
    i : INT;
END_VAR
_M_CopySet := FALSE;
_exportNext := 0;
IF _configStore = 0 THEN RETURN; END_IF
IF NOT _configStore.M_ReadInfo(SetName := SetName, Info := info) THEN RETURN; END_IF
IF (info.SetName <> SetName) OR (info.RecordCount < 1)
OR (info.RecordCount > PL_Fraktal.MAX_SET_RECORDS) THEN RETURN; END_IF
IF NOT _loadSnapshot.M_SaveBegin(Info := info) THEN RETURN; END_IF
FOR i := 1 TO info.RecordCount DO
    IF NOT _configStore.M_ReadRecord(SetName := SetName, Index := i, Record := record) THEN
        _loadSnapshot.M_SaveAbort(); RETURN;
    END_IF
    IF NOT _loadSnapshot.M_SaveRecord(Record := record) THEN
        _loadSnapshot.M_SaveAbort(); RETURN;
    END_IF
END_FOR
_M_CopySet := _loadSnapshot.M_SaveCommit();
END_METHOD

// Reuse the capability walk for immutable export and complete-set validation.
METHOD PRIVATE _M_CaptureConfig : BOOL
VAR_INPUT
    SetName : STRING(80);
    Kind : E_ConfigKind;
    ModelIndex : UDINT;
END_VAR
_exportNext := 0; // every replacement invalidates the old immutable cursor
_M_CaptureConfig := _M_CaptureInto(Store := _snapshot, SetName := SetName, Kind := Kind,
    ModelIndex := ModelIndex);
END_METHOD

// The capability walk as one set in Store. The live documents capture into
// _loadSnapshot, so writing them never invalidates an export of _snapshot.
METHOD PRIVATE _M_CaptureInto : BOOL
VAR_INPUT
    Store : I_ConfigStore;
    SetName : STRING(80);
    Kind : E_ConfigKind;
    ModelIndex : UDINT;
END_VAR
VAR
    info : ST_ConfigSetInfo;
    records : INT;
END_VAR
_M_CaptureInto := FALSE;
IF NOT _M_OpenModelView(Index := ModelIndex) THEN RETURN; END_IF
info.SetName := SetName;
info.Used := TRUE;
info.RootIdentity := Status.Name;
info.SetSchema := CONFIG_SET_SCHEMA;
info.ConfigRev := ConfigRev;
info.Kind := Kind;
info.ModelCode := Model.ModelCode;
IF ModelIndex > 0 THEN info.ModelCode := AvailableModels[ModelIndex].ModelCode; END_IF
IF Kind <> E_ConfigKind.PAR_CFG THEN info.ModelCode := ''; END_IF
info.CreatedAt := F_Now();
info.TimeSynchronized := F_TimeSynchronized();
IF _configPager.M_SetupSetSave(Store := Store, Info := info) THEN
    M_AppendConfig(Pager := _configPager);
    _M_CaptureInto := _configPager.M_FinishSetSave(Records => records);
END_IF
_pModelView := 0;
END_METHOD

